(* IEC 61131-3 sources: plc_NativeGateway/src, 67 files *)

(* ---- NG_Add4.st ---- *)
FUNCTION NG_Add4 : DWORD
VAR_INPUT
    a : DWORD;
    b : DWORD;
    c : DWORD;
    d : DWORD;
END_VAR
(* Four uint32 operands fit uint64. A mask implements modulo 2^32 without
   software uint64 division on the AXC F 2152 ARM target. *)
NG_Add4 := TO_DWORD(TO_LWORD(TO_ULINT(a)+TO_ULINT(b)+TO_ULINT(c)+TO_ULINT(d)) AND LWORD#16#FFFFFFFF);
END_FUNCTION

(* ---- NG_Allowed.st ---- *)
FUNCTION NG_Allowed : BOOL
VAR_INPUT
    Parent : INT;
    Keys : NG_Text; (* Delimited with |, including first and last separator. *)
END_VAR
VAR_INPUT
    Doc : NG_Document;
END_VAR
VAR
    i : INT;
    key : STRING[68];
END_VAR
NG_Allowed := FALSE;
IF (Parent < 1) OR (Parent > Doc.Count) THEN RETURN; END_IF;
IF Doc.Tokens[Parent].Kind <> 1 THEN RETURN; END_IF;
i := Parent + 1;
WHILE i < Doc.Tokens[Parent].NextToken DO
    key := CONCAT('|', Doc.Tokens[i].Key, '|');
    IF FIND(Keys,key) = 0 THEN RETURN; END_IF;
    IF Doc.Tokens[i].NextToken <= i THEN RETURN; END_IF;
    i := Doc.Tokens[i].NextToken;
END_WHILE;
NG_Allowed := TRUE;
END_FUNCTION

(* ---- NG_Bool.st ---- *)
FUNCTION NG_Bool : STRING
VAR_INPUT
    Value : BOOL;
END_VAR
IF Value THEN NG_Bool := 'true'; ELSE NG_Bool := 'false'; END_IF;
END_FUNCTION

(* ---- NG_CheckConfig.st ---- *)
FUNCTION NG_CheckConfig : NG_Text
VAR_INPUT
    Config : NG_Config;
END_VAR
VAR
    d : INT;
    p : INT;
    i : INT;
    width : UDINT;
    point : NG_Point;
END_VAR
NG_CheckConfig := 'SCHEMA_INVALID';
IF (Config.PointCount < 0) OR (Config.PointCount > 320) THEN RETURN; END_IF;
IF (Config.DeviceCount < 0) OR (Config.DeviceCount > 50) OR (Config.batchIntervalMs < 1) OR (Config.batchIntervalMs > 86400000) OR (Config.maxBatchPoints < 1) OR (Config.maxBatchPoints > 500) THEN RETURN; END_IF;
FOR d := 1 TO Config.DeviceCount DO
    IF NOT NG_ValidId(Config.Devices[d].deviceId) THEN RETURN; END_IF;
    FOR i := 1 TO d-1 DO
        IF Config.Devices[d].deviceId = Config.Devices[i].deviceId THEN NG_CheckConfig := 'DUPLICATE_DEVICE_ID'; RETURN; END_IF;
    END_FOR;
    IF NOT NG_IPv4(Config.Devices[d].host) THEN NG_CheckConfig := 'BAD_CONFIGURATION'; RETURN; END_IF;
    IF (Config.Devices[d].port = 0) OR (Config.Devices[d].PointCount < 0) OR (Config.Devices[d].PointCount > 32) THEN RETURN; END_IF;
    IF (Config.Devices[d].connectTimeoutMs < 1) OR (Config.Devices[d].connectTimeoutMs > 300000) OR (Config.Devices[d].requestTimeoutMs < 1) OR (Config.Devices[d].requestTimeoutMs > 300000) OR (Config.Devices[d].retryCount > 10) THEN RETURN; END_IF;
    IF (Config.Devices[d].maxReadRegisters > UINT#125) OR (Config.Devices[d].hasMaxRegisterGap AND (Config.Devices[d].maxRegisterGap > UINT#124)) THEN RETURN; END_IF;
    FOR p := 1 TO Config.Devices[d].PointCount DO
        point := Config.Points[Config.Devices[d].PointStart+p-1];
        IF NOT NG_ValidId(point.pointId) THEN RETURN; END_IF;
        FOR i := 1 TO p-1 DO
            IF point.pointId = Config.Points[Config.Devices[d].PointStart+i-1].pointId THEN NG_CheckConfig := 'DUPLICATE_POINT_ID'; RETURN; END_IF;
        END_FOR;
        IF (point.pollIntervalMs < 1) OR (point.pollIntervalMs > 86400000) OR (point.reportIntervalMs < 1) OR (point.reportIntervalMs > 86400000) OR (point.staleAfterMs > 86400000) OR (point.deadband < 0) THEN RETURN; END_IF;
        IF point.staleAfterMs < point.pollIntervalMs THEN NG_CheckConfig := 'INVALID_STALE_INTERVAL'; RETURN; END_IF;
        IF (point.reportMode <> 'cyclic') AND (point.reportMode <> 'change') AND (point.reportMode <> 'change_or_cyclic') THEN RETURN; END_IF;
        IF point.dataType = 'bool' THEN
            width := 1;
            IF (point.area <> 'coil') AND (point.area <> 'discrete_input') THEN RETURN; END_IF;
            IF (point.byteOrder <> '') OR (point.scale <> 1) OR (point.offset <> 0) OR (point.deadband <> 0) THEN RETURN; END_IF;
        ELSE
            IF (point.area <> 'holding_register') AND (point.area <> 'input_register') THEN RETURN; END_IF;
            IF (point.dataType = 'uint16') OR (point.dataType = 'int16') THEN
                width := 1;
                IF (point.byteOrder <> 'AB') AND (point.byteOrder <> 'BA') THEN RETURN; END_IF;
            ELSIF (point.dataType = 'uint32') OR (point.dataType = 'int32') OR (point.dataType = 'float32') THEN
                width := 2;
                IF (point.byteOrder <> 'ABCD') AND (point.byteOrder <> 'BADC') AND (point.byteOrder <> 'CDAB') AND (point.byteOrder <> 'DCBA') THEN RETURN; END_IF;
            ELSE RETURN;
            END_IF;
        END_IF;
        IF TO_UDINT(point.address) + width > 65536 THEN NG_CheckConfig := 'INVALID_ADDRESS'; RETURN; END_IF;
    END_FOR;
END_FOR;
NG_CheckConfig := '';
END_FUNCTION

(* ---- NG_Clip.st ---- *)
FUNCTION NG_Clip : NG_Text
VAR_INPUT
    Value : NG_Text;
END_VAR
IF LEN(Value) > 48 THEN NG_Clip := CONCAT(LEFT(Value,45),'...');
ELSE NG_Clip := Value; END_IF;
END_FUNCTION

(* ---- NG_IPv4.st ---- *)
FUNCTION NG_IPv4 : BOOL
VAR_INPUT
    Host : STRING[253];
END_VAR
VAR
    i : INT;
    dots : INT;
    digits : INT;
    value : INT;
    c : STRING[1];
END_VAR
NG_IPv4 := FALSE; dots := 0; digits := 0; value := 0;
FOR i := 1 TO LEN(Host) DO
    c := MID(Host,1,i);
    IF c = '.' THEN
        IF (digits = 0) OR (value > 255) THEN RETURN; END_IF;
        dots := dots + 1; digits := 0; value := 0;
    ELSIF (c >= '0') AND (c <= '9') THEN
        value := value * 10 + TO_INT(c); digits := digits + 1;
        IF digits > 3 THEN RETURN; END_IF;
    ELSE RETURN;
    END_IF;
END_FOR;
NG_IPv4 := (dots = 3) AND (digits > 0) AND (value <= 255);
END_FUNCTION

(* ---- NG_Member.st ---- *)
FUNCTION NG_Member : INT
VAR_INPUT
    Parent : INT;
    Key : NG_Id;
END_VAR
VAR_INPUT
    Doc : NG_Document;
END_VAR
VAR
    i : INT;
END_VAR
NG_Member := 0;
IF (Parent < 1) OR (Parent > Doc.Count) THEN RETURN; END_IF;
i := Parent + 1;
WHILE i < Doc.Tokens[Parent].NextToken DO
    IF Doc.Tokens[i].Key = Key THEN NG_Member := i; RETURN; END_IF;
    IF Doc.Tokens[i].NextToken <= i THEN RETURN; END_IF;
    i := Doc.Tokens[i].NextToken;
END_WHILE;
END_FUNCTION

(* ---- NG_NumberValid.st ---- *)
FUNCTION NG_NumberValid : BOOL
VAR_INPUT
    s : NG_Text;
END_VAR
VAR
    i : INT;
    n : INT;
    start : INT;
    c : STRING[1];
END_VAR
NG_NumberValid := FALSE;
n := LEN(s); i := 1;
IF n = 0 THEN RETURN; END_IF;
IF MID(s,1,i) = '-' THEN i := i + 1; END_IF;
IF i > n THEN RETURN; END_IF;
c := MID(s,1,i);
IF c = '0' THEN
    i := i + 1;
ELSIF (c >= '1') AND (c <= '9') THEN
    WHILE i <= n DO
        c := MID(s,1,i);
        IF (c < '0') OR (c > '9') THEN EXIT; END_IF;
        i := i + 1;
    END_WHILE;
ELSE RETURN;
END_IF;
IF i > n THEN NG_NumberValid := TRUE; RETURN; END_IF;
IF MID(s,1,i) = '.' THEN
    i := i + 1; start := i;
    WHILE i <= n DO
        c := MID(s,1,i);
        IF (c < '0') OR (c > '9') THEN EXIT; END_IF;
        i := i + 1;
    END_WHILE;
    IF i = start THEN RETURN; END_IF;
END_IF;
IF i > n THEN NG_NumberValid := TRUE; RETURN; END_IF;
c := MID(s,1,i);
IF (c = 'e') OR (c = 'E') THEN
    i := i + 1; IF i > n THEN RETURN; END_IF; c := MID(s,1,i);
    IF (c = '+') OR (c = '-') THEN i := i + 1; END_IF;
    start := i;
    WHILE i <= n DO
        c := MID(s,1,i);
        IF (c < '0') OR (c > '9') THEN EXIT; END_IF;
        i := i + 1;
    END_WHILE;
    IF i = start THEN RETURN; END_IF;
END_IF;
NG_NumberValid := i = n + 1;
END_FUNCTION

(* ---- NG_ProcNumber.st ---- *)
FUNCTION NG_ProcNumber : ULINT
VAR_INPUT
    Text : NG_ProcText;
    Key : STRING[64];
END_VAR
VAR
    p : INT;
    n : INT;
    c : INT;
    started : BOOL;
END_VAR
NG_ProcNumber := 0; started := FALSE; p := FIND(Text,Key); IF p = 0 THEN RETURN; END_IF;
p := p+LEN(Key); n := LEN(Text);
WHILE p <= n DO
    c := GET_CHAR(Text,p);
    IF (c >= 48) AND (c <= 57) THEN NG_ProcNumber := NG_ProcNumber*10+TO_ULINT(c-48); started := TRUE;
    ELSIF started OR ((c <> 32) AND (c <> 9)) THEN RETURN;
    END_IF;
    p := p+1;
END_WHILE;
END_FUNCTION

(* ---- NG_QualityCode.st ---- *)
FUNCTION NG_QualityCode : USINT
VAR_INPUT
    Quality : STRING[24];
END_VAR
NG_QualityCode := 7;
IF Quality='UNKNOWN' THEN NG_QualityCode:=1;
ELSIF Quality='GOOD' THEN NG_QualityCode:=2;
ELSIF Quality='STALE' THEN NG_QualityCode:=3;
ELSIF Quality='BAD_CONNECTION' THEN NG_QualityCode:=4;
ELSIF Quality='BAD_TIMEOUT' THEN NG_QualityCode:=5;
ELSIF Quality='BAD_PROTOCOL' THEN NG_QualityCode:=6;
END_IF;
END_FUNCTION

(* ---- NG_QualityName.st ---- *)
FUNCTION NG_QualityName : NG_Text
VAR_INPUT
    Code : USINT;
END_VAR
CASE Code OF
2: NG_QualityName:='GOOD';
3: NG_QualityName:='STALE';
4: NG_QualityName:='BAD_CONNECTION';
5: NG_QualityName:='BAD_TIMEOUT';
6: NG_QualityName:='BAD_PROTOCOL';
7: NG_QualityName:='BAD_DECODE';
ELSE NG_QualityName:='UNKNOWN';
END_CASE;
END_FUNCTION

(* ---- NG_Quote.st ---- *)
FUNCTION NG_Quote : NG_Quoted
VAR_INPUT
    s : NG_Text;
END_VAR
VAR
    i : INT;
    c : STRING[1];
    character : INT;
    plain : BOOL;
    characters : ARRAY[0..255] OF BYTE;
    copied : BOOL;
    length : INT;
END_VAR
(* Scan once for escaping; common identities take one final concatenation. *)
plain:=TRUE;
length:=LEN(s); copied:=TRUE;
IF length>0 THEN copied:=STRING_COPY(s,characters,UDINT#0,TO_UDINT(length)); END_IF;
FOR i:=1 TO length DO
    IF copied THEN character:=TO_INT(characters[i-1]);
    ELSE character:=GET_CHAR(s,i); END_IF;
    IF (character<32) OR (character=34) OR (character=92) THEN plain:=FALSE; EXIT; END_IF;
END_FOR;
IF plain THEN NG_Quote:=CONCAT('"',s,'"'); RETURN; END_IF;
NG_Quote := '"';
FOR i := 1 TO LEN(s) DO
    c := MID(s,1,i);
    IF c = '"' THEN NG_Quote := CONCAT(NG_Quote,'\\','"');
    ELSIF c = '\\' THEN NG_Quote := CONCAT(NG_Quote,'\\\\');
    ELSIF c = '\n' THEN NG_Quote := CONCAT(NG_Quote,'\\n');
    ELSIF GET_CHAR(c,1) = 13 THEN NG_Quote := CONCAT(NG_Quote,'\\r');
    ELSIF c = '\t' THEN NG_Quote := CONCAT(NG_Quote,'\\t');
    ELSE NG_Quote := CONCAT(NG_Quote,c);
    END_IF;
END_FOR;
NG_Quote := CONCAT(NG_Quote,'"');
END_FUNCTION

(* ---- NG_Range.st ---- *)
FUNCTION NG_Range : BOOL
VAR_INPUT
    Text : NG_Text;
    Minimum : LREAL;
    Maximum : LREAL;
    IntegerOnly : BOOL;
END_VAR
VAR
    n : LREAL;
END_VAR
NG_Range := FALSE;
IF NOT NG_NumberValid(Text) OR (LEN(Text)>20) THEN RETURN; END_IF;
(* UI configuration values do not need exponent notation. *)
IF (FIND(Text,'e')>0) OR (FIND(Text,'E')>0) THEN RETURN; END_IF;
n := TO_LREAL(Text);
NG_Range := (n >= Minimum) AND (n <= Maximum);
IF IntegerOnly AND (n <> TO_LREAL(TO_LINT(n))) THEN NG_Range := FALSE; END_IF;
END_FUNCTION

(* ---- NG_SafeAdd.st ---- *)
FUNCTION NG_SafeAdd : ULINT
VAR_INPUT
    CounterValue : ULINT;
    Delta : ULINT;
END_VAR
IF CounterValue>=ULINT#9007199254740991 THEN NG_SafeAdd:=ULINT#9007199254740991; RETURN; END_IF;
IF Delta>ULINT#9007199254740991-CounterValue THEN
    NG_SafeAdd := ULINT#9007199254740991;
ELSE NG_SafeAdd := CounterValue+Delta;
END_IF;
END_FUNCTION

(* ---- NG_UiJoin.st ---- *)
FUNCTION NG_UiJoin : NG_UiLabel
VAR_INPUT
    A : NG_UiLabel;
    B : NG_UiLabel;
    C : NG_UiLabel;
    D : NG_UiLabel;
    E : NG_UiLabel;
    F : NG_UiLabel;
    G : NG_UiLabel;
    H : NG_UiLabel;
END_VAR
VAR
    Buffer : NG_UiLabel;
    Parts : ARRAY[1..8] OF NG_UiLabel;
    Chunk : NG_UiLabel;
    Remaining : INT;
    i : INT;
END_VAR
(* Explicit intermediates avoid the vendor's default 80-character FU temporary. *)
Parts[1]:=A; Parts[2]:=B; Parts[3]:=C; Parts[4]:=D;
Parts[5]:=E; Parts[6]:=F; Parts[7]:=G; Parts[8]:=H;
Buffer:="";
FOR i:=1 TO 8 DO
    Remaining:=256-LEN(Buffer);
    IF Remaining<=0 THEN EXIT; END_IF;
    Chunk:=Parts[i];
    IF LEN(Chunk)>Remaining THEN Chunk:=LEFT_WSTRING(Chunk,Remaining); END_IF;
    Buffer:=CONCAT_WSTRING(Buffer,Chunk);
END_FOR;
NG_UiJoin:=Buffer;
END_FUNCTION

(* ---- NG_UiText.st ---- *)
FUNCTION NG_UiText : NG_UiLabel
VAR_INPUT
    Value : NG_Text;
    English : BOOL;
END_VAR
NG_UiText:=TO_WSTRING(Value,"");
IF English THEN
IF Value='PERSISTED' THEN NG_UiText:="Saved · no changes";
ELSIF Value='UNSAVED DRAFT' THEN NG_UiText:="Unapplied changes";
ELSIF Value='VERSION CONFLICT' THEN NG_UiText:="Configuration changed";
ELSIF Value='CONNECTED' THEN NG_UiText:="Connected";
ELSIF Value='CONNECTING' THEN NG_UiText:="Connecting";
ELSIF Value='HUB_MANAGED' THEN NG_UiText:="Hub managed";
ELSIF Value='STANDALONE' THEN NG_UiText:="Local maintenance";
ELSIF Value='holding_register' THEN NG_UiText:="Holding register";
ELSIF Value='input_register' THEN NG_UiText:="Input register";
ELSIF Value='discrete_input' THEN NG_UiText:="Discrete input";
ELSIF Value='cyclic' THEN NG_UiText:="Cyclic";
ELSIF Value='change' THEN NG_UiText:="On change";
ELSIF Value='change_or_cyclic' THEN NG_UiText:="Change or cyclic";
ELSIF Value='Startup identity persisted; MQTT starting.' THEN NG_UiText:="Saved configuration restored automatically. No need to save again.";
ELSIF Value='true' THEN NG_UiText:="Enabled";
ELSIF Value='TRUE' THEN NG_UiText:="Enabled";
ELSIF Value='false' THEN NG_UiText:="Disabled";
ELSIF Value='FALSE' THEN NG_UiText:="Disabled";
ELSIF Value='HUB_MANAGED - local device/point changes blocked' THEN NG_UiText:="Managed by Hub: edit and publish devices, points and periods in Hub. Connection maintenance is available here.";
ELSIF Value='STANDALONE - local maintenance enabled' THEN NG_UiText:="Standalone: edit devices and points → save to draft → review and activate.";
END_IF;
RETURN;
END_IF;
IF Value='Open the management mode confirmation before saving.' THEN NG_UiText:="请先打开模式切换确认页，检查选项后再确认。";
ELSIF Value='Waiting for initial Hub configuration. Existing local acquisition is retained.' THEN NG_UiText:="正在等待平台首次配置；现有本地采集保留，暂不向平台上报。";
ELSIF Value='Invalid management mode.' THEN NG_UiText:="管理模式无效，请重新选择平台管理或本地维护。";
ELSIF Value='MAINTENANCE - incoming platform configuration locked' THEN NG_UiText:="本地维护：平台配置暂不应用；修改后请交还平台，避免两端配置冲突。";
ELSIF Value='Hub owns configuration. Local maintenance requires manual confirmation.' THEN NG_UiText:="当前由平台管理。需要本地编辑时，请手动进入维护。";
ELSIF Value='Local changes active. Acquisition continues; Hub data reporting is paused.' THEN NG_UiText:="本地改动已生效：继续采集，暂停写入平台；交还时恢复平台配置。";
ELSIF Value='Local maintenance active. Hub configuration is locked until you return ownership.' THEN NG_UiText:="本地维护中：平台配置暂不应用。维护完成后请交还平台。";
ELSIF Value='The selected management mode is already active.' THEN NG_UiText:="已处于所选模式，无需重复切换。";
ELSIF Value='Saving management mode; existing identity is retained.' THEN NG_UiText:="正在保存管理模式，保留当前网关标识。";
ELSIF Value='Management mode saved. Check the ownership guidance above.' THEN NG_UiText:="管理模式已保存并生效，请查看上方的管理说明。";
ELSIF Value='Clearing local configuration and version baseline...' THEN NG_UiText:="正在清空本地点表与版本基线，请稍候。";
ELSIF Value='Open the reset confirmation before clearing local configuration.' THEN NG_UiText:="请先打开重置确认页后再确认清空。";
ELSIF Value='Local configuration and version baseline cleared; requesting fresh config from Hub.' THEN NG_UiText:="已清空本地点表与版本基线，正在重连并向平台重新拉取配置。";
ELSIF Value='Check broker URI, gateway ID, client ID and time zone.' THEN NG_UiText:="请检查服务器地址、网关标识与时区。";
ELSIF Value='Broker settings saved; configuration ownership is unchanged.' THEN NG_UiText:="连接设置已保存，正在重连；管理模式保持不变。";
ELSIF Value='CONNECTED' THEN NG_UiText:="已连接";
ELSIF Value='CONNECTING' THEN NG_UiText:="正在连接";
ELSIF Value='ONLINE' THEN NG_UiText:="在线";
ELSIF Value='OFFLINE' THEN NG_UiText:="离线";
ELSIF Value='DEGRADED' THEN NG_UiText:="部分异常";
ELSIF Value='DISABLED' THEN NG_UiText:="已停用";
ELSIF Value='UNCONFIGURED' THEN NG_UiText:="未配置";
ELSIF Value='DRAFT' THEN NG_UiText:="待生效";
ELSIF Value='GOOD' THEN NG_UiText:="正常";
ELSIF Value='BAD' THEN NG_UiText:="异常";
ELSIF Value='STALE' THEN NG_UiText:="已过期";
ELSIF Value='UNKNOWN' THEN NG_UiText:="暂无数据";
ELSIF Value='BAD_COMMUNICATION' THEN NG_UiText:="通信异常";
ELSIF Value='BAD_CONFIGURATION' THEN NG_UiText:="配置有误";
ELSIF Value='true' THEN NG_UiText:="启用";
ELSIF Value='TRUE' THEN NG_UiText:="启用";
ELSIF Value='false' THEN NG_UiText:="停用";
ELSIF Value='FALSE' THEN NG_UiText:="停用";
ELSIF Value='PERSISTED' THEN NG_UiText:="已保存，无待生效修改";
ELSIF Value='UNSAVED DRAFT' THEN NG_UiText:="有待生效的修改";
ELSIF Value='VERSION CONFLICT' THEN NG_UiText:="配置已变更，请放弃旧草稿";
ELSIF Value='HUB_MANAGED' THEN NG_UiText:="平台统一管理";
ELSIF Value='STANDALONE' THEN NG_UiText:="本地维护";
ELSIF Value='HUB_MANAGED - local device/point changes blocked' THEN NG_UiText:="平台管理：在 Hub 编辑设备、点位与周期并发布；此处查看和维护连接。";
ELSIF Value='STANDALONE - local maintenance enabled' THEN NG_UiText:="本地管理：编辑设备和点位 → 保存到待生效配置 → 确认生效并保存。";
ELSIF Value='holding_register' THEN NG_UiText:="保持寄存器";
ELSIF Value='input_register' THEN NG_UiText:="输入寄存器";
ELSIF Value='coil' THEN NG_UiText:="线圈";
ELSIF Value='discrete_input' THEN NG_UiText:="离散输入";
ELSIF Value='cyclic' THEN NG_UiText:="定时上报";
ELSIF Value='change' THEN NG_UiText:="变化时上报";
ELSIF Value='change_or_cyclic' THEN NG_UiText:="变化或定时上报";
ELSIF Value='voltage' THEN NG_UiText:="电压";
ELSIF Value='current' THEN NG_UiText:="电流";
ELSIF Value='frequency' THEN NG_UiText:="频率";
ELSIF Value='power' THEN NG_UiText:="功率";
ELSIF Value='energy' THEN NG_UiText:="累计电能";
ELSIF Value='No device selected' THEN NG_UiText:="暂无设备，请先添加设备";
ELSIF Value='No point selected' THEN NG_UiText:="暂无点位，请先添加点位";
ELSIF Value='HUB_MANAGED: publish device and point changes from Hub.' THEN NG_UiText:="当前由平台管理，请在 Hub 修改并发布设备和点位配置。";
ELSIF Value='Display refreshed from active configuration. Unapplied draft discarded.' THEN NG_UiText:="已按当前运行配置更新显示，未生效的草稿已放弃。";
ELSIF Value='Loaded persisted active configuration.' THEN NG_UiText:="已按控制器当前运行配置更新显示。";
ELSIF Value='Capacity reached: 50 devices.' THEN NG_UiText:="设备数量已达上限：50 台。";
ELSIF Value='Capacity reached: 32 points/device, 320 shared points.' THEN NG_UiText:="点位数量已达上限：每台 32 个，总计 320 个。";
ELSIF Value='New device: save into draft, then add its points.' THEN NG_UiText:="填写连接参数并保存设备，再为该设备添加点位。";
ELSIF Value='Save a device into the draft first.' THEN NG_UiText:="请先保存设备，再添加该设备的点位。";
ELSIF Value='New point: save into draft, then apply the complete draft.' THEN NG_UiText:="填写寄存器与周期，保存点位后再确认配置生效。";
ELSIF Value='Busy: configuration transaction in progress. Try again shortly.' THEN NG_UiText:="正在保存配置，请稍候再试。";
ELSIF Value='Device index 1..50; point index 1..32.' THEN NG_UiText:="请检查设备序号（1～50）和点位序号（1～32）。";
ELSIF Value='Invalid device fields: check ID, name, IPv4, port and timeout values.' THEN NG_UiText:="设备未保存：检查唯一标识、名称、地址、端口与超时。";
ELSIF Value='Device saved to draft. Apply draft to persist.' THEN NG_UiText:="设备已加入待生效配置。检查点位后，点击“使配置生效”。";
ELSIF Value='Invalid point fields; save the device first and check numeric fields.' THEN NG_UiText:="点位未保存：先保存设备，再检查地址、周期、倍率等数值。";
ELSIF Value='Point saved to draft. Apply draft to persist.' THEN NG_UiText:="点位已加入待生效配置。点击“使配置生效”后开始使用。";
ELSIF Value='Device and points removed from draft. Apply to persist.' THEN NG_UiText:="设备及其点位已从草稿移除，确认配置生效后才停止采集。";
ELSIF Value='Point removed from draft. Apply to persist.' THEN NG_UiText:="点位已从草稿移除，确认配置生效后才停止采集。";
ELSIF Value='Invalid device polling/report period.' THEN NG_UiText:="周期未修改：采集与上报周期必须为有效的毫秒数。";
ELSIF Value='Device point periods updated in draft. Apply to persist.' THEN NG_UiText:="该设备的点位周期已加入待生效配置，请确认生效。";
ELSIF Value='VERSION_CONFLICT: reload active configuration before applying.' THEN NG_UiText:="运行配置已有更新。请放弃旧草稿，按最新配置重新编辑。";
ELSIF Value='Invalid gateway batch settings.' THEN NG_UiText:="请检查组批周期与每包点数（1～64）。";
ELSIF Value='Saving, hashing and reading back configuration...' THEN NG_UiText:="正在保存并校验配置，请稍候。";
ELSIF Value='Check broker/mode/ID. Mode change requires a new Gateway ID to isolate configuration history.' THEN NG_UiText:="连接未保存：检查地址、网关标识、客户端标识与模式；换模式须换网关标识。";
ELSIF Value='Saving broker settings...' THEN NG_UiText:="正在保存消息服务器连接设置，请稍候。";
ELSIF Value='APPLIED: configuration saved and activated.' THEN NG_UiText:="配置已生效并保存；重启后将自动恢复。";
ELSIF Value='Broker/mode saved; identity changes reset local baseline.' THEN NG_UiText:="连接设置已保存，正在自动重连；新身份需由平台重新下发配置。";
ELSIF Value='Startup identity persisted; MQTT starting.' THEN NG_UiText:="已自动恢复保存的配置，无需重复保存。";
ELSIF Value='Persisting unique startup identity before MQTT...' THEN NG_UiText:="正在保存启动信息，随后自动连接消息服务器。";
ELSIF Value='STORAGE_ERROR: active configuration unchanged.' THEN NG_UiText:="保存失败，运行配置保持原样。请检查控制器存储。";
ELSIF Value='Saving / validating durable file...' THEN NG_UiText:="正在写入并校验控制器配置文件……";
ELSIF Value='STORAGE ERROR: configuration not committed.' THEN NG_UiText:="配置保存失败，请检查控制器存储。";
ELSIF Value='Restoring saved configuration...' THEN NG_UiText:="正在恢复已保存配置，随后自动连接并采集。";
ELSIF Value='Broker unavailable. Retrying automatically; local acquisition continues.' THEN NG_UiText:="消息服务器暂不可用，正在自动重连；本地采集继续运行。";
ELSIF Value='MQTT_DISCONNECTED' THEN NG_UiText:="连接中断，自动重连中";
ELSIF Value='MQTT_CONNECT_ERROR' THEN NG_UiText:="连接失败，自动重试中";
ELSIF Value='MQTT_TIMEOUT' THEN NG_UiText:="连接超时，自动重试中";
ELSIF Value='MQTT_PUBLISH_ERROR' THEN NG_UiText:="发送失败，自动重连中";
ELSIF Value='MQTT_CLIENT_ERROR' THEN NG_UiText:="通信组件异常，自动重试中";
ELSIF Value='MQTT_SUBSCRIBE_ERROR' THEN NG_UiText:="订阅失败，自动重试中";
ELSIF Value='MQTT_CONSUME_ERROR' THEN NG_UiText:="接收失败，自动重试中";
ELSIF Value='SCHEMA_INVALID' THEN NG_UiText:="配置格式或取值不正确，请检查点位详情。";
ELSIF Value='DUPLICATE_DEVICE_ID' THEN NG_UiText:="设备标识重复，请使用唯一标识。";
ELSIF Value='DUPLICATE_POINT_ID' THEN NG_UiText:="同一设备内点位标识重复。";
ELSIF Value='INVALID_STALE_INTERVAL' THEN NG_UiText:="过期时间必须不小于采集周期。";
ELSIF Value='INVALID_ADDRESS' THEN NG_UiText:="寄存器地址范围无效。";
ELSIF Value='BAD_CONNECTION' THEN NG_UiText:="连接异常";
ELSIF Value='BAD_TIMEOUT' THEN NG_UiText:="请求超时";
ELSIF Value='BAD_PROTOCOL' THEN NG_UiText:="报文异常";
ELSIF Value='BAD_DECODE' THEN NG_UiText:="数据解码异常";
END_IF;
END_FUNCTION

(* ---- NG_Unix.st ---- *)
FUNCTION NG_Unix : ULINT
VAR_INPUT
    Clock : RTC_TYPE;
    UtcOffsetMinutes : INT;
END_VAR
VAR
    y : DINT;
    m : DINT;
    days : LINT;
    md : DINT;
    seconds : LINT;
END_VAR
NG_Unix := 0;
IF (Clock.YEAR < 2020) OR (Clock.YEAR > 2199) OR (Clock.MONTH < 1) OR (Clock.MONTH > 12) OR (Clock.DAY < 1) OR (Clock.DAY > 31) THEN RETURN; END_IF;
days := 0;
FOR y := 1970 TO TO_DINT(Clock.YEAR)-1 DO
    days := days + 365;
    IF ((y MOD 4 = 0) AND (y MOD 100 <> 0)) OR (y MOD 400 = 0) THEN days := days + 1; END_IF;
END_FOR;
FOR m := 1 TO TO_DINT(Clock.MONTH)-1 DO
    CASE m OF
        4,6,9,11: md := 30;
        2:
            md := 28; y := TO_DINT(Clock.YEAR);
            IF ((y MOD 4 = 0) AND (y MOD 100 <> 0)) OR (y MOD 400 = 0) THEN md := 29; END_IF;
        ELSE md := 31;
    END_CASE;
    days := days + md;
END_FOR;
days := days + Clock.DAY - 1;
seconds := days * 86400 + TO_LINT(Clock.HOURS) * 3600 + TO_LINT(Clock.MINUTES) * 60 + Clock.SECONDS - TO_LINT(UtcOffsetMinutes)*60;
IF seconds > 0 THEN NG_Unix := TO_ULINT(seconds)*1000; END_IF;
END_FUNCTION

(* ---- NG_ValidId.st ---- *)
FUNCTION NG_ValidId : BOOL
VAR_INPUT
    s : NG_Id;
END_VAR
VAR
    i : INT;
    c : STRING[1];
END_VAR
NG_ValidId := (LEN(s) > 0) AND (LEN(s) <= 64);
FOR i := 1 TO LEN(s) DO
    c := MID(s, 1, i);
    IF NOT (((c >= 'A') AND (c <= 'Z')) OR ((c >= 'a') AND (c <= 'z')) OR ((c >= '0') AND (c <= '9')) OR ((i > 1) AND ((c = '.') OR (c = '_') OR (c = '-')))) THEN
        NG_ValidId := FALSE;
    END_IF;
END_FOR;
END_FUNCTION

(* ---- NG_WireCode.st ---- *)
FUNCTION NG_WireCode : NG_Text
VAR_INPUT
    Code : NG_Text;
    IsPatch : BOOL;
END_VAR
IF FIND('|SCHEMA_INVALID|INVALID_JSON|PAYLOAD_TOO_LARGE|GATEWAY_MISMATCH|DUPLICATE_DEVICE_ID|DUPLICATE_POINT_ID|DUPLICATE_NODE_ID|INVALID_ADDRESS|INVALID_STALE_INTERVAL|POINT_LIMIT_EXCEEDED|VERSION_CONFLICT|STALE_VERSION|RESOURCE_LIMIT|STORAGE_ERROR|APPLY_FAILED|UNKNOWN_CONFIG_VERSION|UNKNOWN_DEVICE|UNKNOWN_POINT|EXPIRED_DATA|INVALID_TIMESTAMP|DUPLICATE_VALUE|',CONCAT('|',Code,'|')) > 0 THEN NG_WireCode := Code;
ELSIF IsPatch AND (Code = 'RETAINED_PATCH') THEN NG_WireCode := 'OPERATION_CONFLICT';
ELSIF IsPatch AND (FIND('|BASE_CONFIG_MISMATCH|DEVICE_EXISTS|DEVICE_NOT_FOUND|OPERATION_CONFLICT|',CONCAT('|',Code,'|'))>0) THEN NG_WireCode := Code;
ELSE NG_WireCode := 'APPLY_FAILED';
END_IF;
END_FUNCTION

(* ---- NG_AckFields.st ---- *)
FUNCTION_BLOCK NG_AckFields
VAR_INPUT
    Parent : INT;
    ErrorObject : BOOL;
END_VAR
VAR_IN_OUT
    Doc : NG_Document;
END_VAR
VAR_OUTPUT
    Valid : BOOL;
    Fields : ARRAY[1..6] OF INT;
END_VAR
VAR
    i : INT;
    j : INT;
    field : INT;
    count : INT;
END_VAR
(* A bounded, reference-based index for the two ACK object shapes. It keeps
   the full document out of FUNCTION VAR_INPUT argument copies. *)
Valid:=FALSE; FOR j:=1 TO 6 DO Fields[j]:=0; END_FOR;
IF (Parent<1) OR (Parent>Doc.Count) THEN RETURN; END_IF;
IF Doc.Tokens[Parent].Kind<>1 THEN RETURN; END_IF;
i:=Parent+1; count:=0;
WHILE i<Doc.Tokens[Parent].NextToken DO
    count:=count+1; IF count>6 THEN RETURN; END_IF;
    IF (i>Doc.Count) OR (i>8192) THEN RETURN; END_IF;
    field:=0;
    IF ErrorObject THEN
        IF Doc.Tokens[i].Key='code' THEN field:=1;
        ELSIF Doc.Tokens[i].Key='path' THEN field:=2;
        ELSIF Doc.Tokens[i].Key='message' THEN field:=3;
        ELSIF Doc.Tokens[i].Key='deviceId' THEN field:=4;
        ELSIF Doc.Tokens[i].Key='pointId' THEN field:=5; END_IF;
    ELSE
        IF Doc.Tokens[i].Key='schemaVersion' THEN field:=1;
        ELSIF Doc.Tokens[i].Key='gatewayId' THEN field:=2;
        ELSIF Doc.Tokens[i].Key='timestamp' THEN field:=3;
        ELSIF Doc.Tokens[i].Key='messageId' THEN field:=4;
        ELSIF Doc.Tokens[i].Key='status' THEN field:=5;
        ELSIF Doc.Tokens[i].Key='errors' THEN field:=6; END_IF;
    END_IF;
    IF field=0 THEN RETURN; END_IF;
    IF Fields[field]<>0 THEN RETURN; END_IF;
    Fields[field]:=i;
    IF (Doc.Tokens[i].NextToken<=i) OR (Doc.Tokens[i].NextToken>Doc.Tokens[Parent].NextToken) THEN RETURN; END_IF;
    i:=Doc.Tokens[i].NextToken;
END_WHILE;
IF i<>Doc.Tokens[Parent].NextToken THEN RETURN; END_IF;
IF ErrorObject THEN
    IF (Fields[1]=0) OR (Fields[2]=0) OR (Fields[3]=0) THEN RETURN; END_IF;
ELSE
    FOR j:=1 TO 6 DO IF Fields[j]=0 THEN RETURN; END_IF; END_FOR;
END_IF;
Valid:=TRUE;
END_FUNCTION_BLOCK

(* ---- NG_AuditAssociation.st ---- *)
FUNCTION_BLOCK NG_AuditAssociation
VAR_INPUT
    Slot : UINT;
    MessageId : NG_Id;
END_VAR
VAR_IN_OUT
    Buffer : NG_Buffer;
END_VAR
VAR
    index : UINT;
    configSlot : UINT;
    j : UINT;
    offset : UINT;
END_VAR
IF NOT Buffer.AuditEnabled THEN RETURN; END_IF;
IF (Slot<1) OR (Slot>16) THEN Buffer.CaptureStopped:=TRUE; Buffer.EvidenceComplete:=FALSE; RETURN; END_IF;
IF Buffer.AssociationWriteSeq>=ULINT#9007199254740991 THEN Buffer.CaptureStopped:=TRUE; RETURN; END_IF;
IF Buffer.AssociationWriteSeq-Buffer.AssociationReadSeq>=32 THEN
    index:=TO_UINT(Buffer.AssociationReadSeq MOD 32)+1;
    configSlot:=Buffer.Associations[index].ConfigSlot;
    IF (configSlot<1) OR (configSlot>4) THEN Buffer.CaptureStopped:=TRUE; Buffer.EvidenceComplete:=FALSE; RETURN; END_IF;
    IF Buffer.Configs[configSlot].References=0 THEN Buffer.CaptureStopped:=TRUE; Buffer.EvidenceComplete:=FALSE; RETURN; END_IF;
    Buffer.Configs[configSlot].References:=Buffer.Configs[configSlot].References-1;
    Buffer.AssociationReadSeq:=Buffer.AssociationReadSeq+1;
    Buffer.AssociationDropped:=NG_SafeAdd(Buffer.AssociationDropped,ULINT#1); Buffer.EvidenceComplete:=FALSE;
END_IF;
Buffer.AssociationWriteSeq:=Buffer.AssociationWriteSeq+1; index:=TO_UINT((Buffer.AssociationWriteSeq-1) MOD 32)+1;
configSlot:=Buffer.BatchOwners[Slot].ConfigSlot;
IF (configSlot<1) OR (configSlot>4) THEN Buffer.CaptureStopped:=TRUE; Buffer.EvidenceComplete:=FALSE; RETURN; END_IF;
Buffer.Associations[index].Ordinal:=Buffer.AssociationWriteSeq;
Buffer.Associations[index].MessageId:=MessageId; Buffer.Associations[index].Digest:=Buffer.BatchOwners[Slot].Digest;
Buffer.Associations[index].ConfigSlot:=configSlot; Buffer.Associations[index].ConfigGeneration:=Buffer.Configs[configSlot].Generation;
Buffer.Associations[index].BatchGeneration:=Buffer.BatchGenerations[Slot]; Buffer.Associations[index].Category:=Buffer.BatchOwners[Slot].Category;
Buffer.Associations[index].Count:=Buffer.BatchOwners[Slot].Count; offset:=(Slot-1)*64;
FOR j:=1 TO Buffer.BatchOwners[Slot].Count DO Buffer.Associations[index].SampleSeqs[j]:=Buffer.Records[Buffer.BatchRefs[offset+j]].SampleSeq; END_FOR;
Buffer.Configs[configSlot].References:=Buffer.Configs[configSlot].References+1;
END_FUNCTION_BLOCK

(* ---- NG_AuditCapture.st ---- *)
FUNCTION_BLOCK NG_AuditCapture
VAR_IN_OUT
    Buffer : NG_Buffer;
    Event : NG_CaptureEvent;
END_VAR
VAR
    index : UINT;
    oldIndex : UINT;
    configSlot : UINT;
END_VAR

IF NOT Buffer.AuditEnabled THEN RETURN; END_IF;
IF (Event.SampleSeq=0) OR (Event.ConfigSlot<1) OR (Event.ConfigSlot>4) THEN
    Buffer.CaptureStopped:=TRUE; Buffer.EvidenceComplete:=FALSE; RETURN;
END_IF;
IF Buffer.AuditWriteSeq-Buffer.AuditReadSeq>=512 THEN
    oldIndex:=TO_UINT(Buffer.AuditReadSeq MOD 512)+1;
    configSlot:=Buffer.AuditEvents[oldIndex].Event.ConfigSlot;
    IF (configSlot<1) OR (configSlot>4) THEN Buffer.CaptureStopped:=TRUE; Buffer.EvidenceComplete:=FALSE; RETURN; END_IF;
    IF Buffer.Configs[configSlot].References=0 THEN Buffer.CaptureStopped:=TRUE; Buffer.EvidenceComplete:=FALSE; RETURN; END_IF;
    Buffer.Configs[configSlot].References:=Buffer.Configs[configSlot].References-1;
    Buffer.AuditReadSeq:=Buffer.AuditReadSeq+1;
    Buffer.AuditDropped:=NG_SafeAdd(Buffer.AuditDropped,ULINT#1); Buffer.EvidenceComplete:=FALSE;
END_IF;
index:=TO_UINT((Event.SampleSeq-1) MOD 512)+1;
Buffer.AuditEvents[index].Event:=Event; Buffer.AuditEvents[index].Decision:=0; Buffer.AuditEvents[index].Reason:=0;
Buffer.Configs[Event.ConfigSlot].References:=Buffer.Configs[Event.ConfigSlot].References+1;
Buffer.AuditWriteSeq:=Event.SampleSeq;
END_FUNCTION_BLOCK

(* ---- NG_AuditDecision.st ---- *)
FUNCTION_BLOCK NG_AuditDecision
VAR_INPUT
    SampleSeq : ULINT;
    Decision : USINT;
    Reason : USINT;
END_VAR
VAR_IN_OUT
    Buffer : NG_Buffer;
END_VAR
VAR
    index : UINT;
END_VAR

IF NOT Buffer.AuditEnabled OR (SampleSeq=0) THEN RETURN; END_IF;
index:=TO_UINT((SampleSeq-1) MOD 512)+1;
IF (SampleSeq>Buffer.AuditReadSeq) AND (Buffer.AuditEvents[index].Event.SampleSeq=SampleSeq) THEN
    Buffer.AuditEvents[index].Decision:=Decision; Buffer.AuditEvents[index].Reason:=Reason;
ELSE Buffer.EvidenceComplete:=FALSE;
END_IF;
END_FUNCTION_BLOCK

(* ---- NG_AuditDrain.st ---- *)
FUNCTION_BLOCK NG_AuditDrain
VAR_INPUT
    BootId : NG_Id;
END_VAR
VAR_IN_OUT
    Buffer : NG_Buffer;
END_VAR
VAR
    index : UINT;
    configSlot : UINT;
    n : INT;
END_VAR
IF (Buffer.AuditAckBootId=BootId) AND (Buffer.AuditAckSeq<=Buffer.AuditWriteSeq) THEN
    FOR n:=1 TO 8 DO
        IF Buffer.AuditReadSeq>=Buffer.AuditAckSeq THEN EXIT; END_IF;
        index:=TO_UINT(Buffer.AuditReadSeq MOD 512)+1;
        IF Buffer.AuditEvents[index].Event.SampleSeq<>Buffer.AuditReadSeq+1 THEN Buffer.EvidenceComplete:=FALSE; RETURN; END_IF;
        IF Buffer.AuditEvents[index].Decision=0 THEN EXIT; END_IF;
        configSlot:=Buffer.AuditEvents[index].Event.ConfigSlot;
        IF (configSlot<1) OR (configSlot>4) THEN Buffer.EvidenceComplete:=FALSE; RETURN; END_IF;
        IF Buffer.Configs[configSlot].References=0 THEN Buffer.EvidenceComplete:=FALSE; RETURN; END_IF;
        Buffer.Configs[configSlot].References:=Buffer.Configs[configSlot].References-1;
        Buffer.AuditReadSeq:=Buffer.AuditReadSeq+1;
    END_FOR;
END_IF;
IF (Buffer.AssociationAckBootId=BootId) AND (Buffer.AssociationAckSeq<=Buffer.AssociationWriteSeq) THEN
    FOR n:=1 TO 4 DO
        IF Buffer.AssociationReadSeq>=Buffer.AssociationAckSeq THEN EXIT; END_IF;
        index:=TO_UINT(Buffer.AssociationReadSeq MOD 32)+1;
        IF Buffer.Associations[index].Ordinal<>Buffer.AssociationReadSeq+1 THEN Buffer.EvidenceComplete:=FALSE; RETURN; END_IF;
        configSlot:=Buffer.Associations[index].ConfigSlot;
        IF (configSlot<1) OR (configSlot>4) THEN Buffer.EvidenceComplete:=FALSE; RETURN; END_IF;
        IF Buffer.Configs[configSlot].References=0 THEN Buffer.EvidenceComplete:=FALSE; RETURN; END_IF;
        Buffer.Configs[configSlot].References:=Buffer.Configs[configSlot].References-1;
        Buffer.AssociationReadSeq:=Buffer.AssociationReadSeq+1;
    END_FOR;
END_IF;
END_FUNCTION_BLOCK

(* ---- NG_BatchBuilder.st ---- *)
FUNCTION_BLOCK NG_BatchBuilder
VAR_INPUT
    GateOpen : BOOL;
    NowMs : ULINT;
    UnixMs : ULINT;
    GatewayId : NG_Id;
    BootId : NG_Id;
    BatchIntervalMs : UDINT;
END_VAR
VAR_IN_OUT
    Buffer : NG_Buffer;
    Packets : ARRAY[1..16] OF NG_Packet;
    Sequence : ULINT;
END_VAR
VAR_OUTPUT
    Busy : BOOL;
END_VAR
VAR
    Digest : NG_StringSHA256;
    Audit : NG_AuditAssociation;
    Stage : UINT;
    Slot : UINT;
    ConfigSlot : UINT;
    Category : UINT;
    q : UINT;
    r : UINT;
    j : UINT;
    offset : UINT;
    countHistory : UINT;
    countNew : UINT;
    n : INT;
    d : INT;
    deviceId : NG_Id;
    valueJson : STRING[80];
    item : STRING[1024];
    bytesNeeded : INT;
    duplicate : BOOL;
    finish : BOOL;
    lastStart : ULINT;
    first : BOOL := TRUE;
    MaterialClockRevision : ULINT;
    windowOpen : BOOL;
    generation : UDINT;
    seenEpoch : UDINT;
    seenPointEpoch : ARRAY[1..320] OF UDINT;
    pointIndex : UINT;
    HeaderUnixMs : ULINT;
    HeaderSequence : ULINT;
    DeviceQuoteSlot : UINT;
    DeviceQuoteGeneration : UDINT;
    DeviceQuoteEpoch : UDINT;
    DeviceQuoteSeen : ARRAY[1..50] OF UDINT;
    DeviceQuotes : ARRAY[1..50] OF STRING[132];
    QuotedDevice : STRING[132];
    ItemPhase : USINT;
    ItemRecord : UINT;
    ItemGeneration : UDINT;
    CachedUtc : ULINT;
    CachedUtcText : STRING[32];
    CachedQuality : USINT;
    CachedQualityText : STRING[40];
    HaveUtc : BOOL;
    HaveQuality : BOOL;
END_VAR
Busy:=Stage<>0;
IF Stage<>0 THEN
    IF (Buffer.BatchGenerations[Slot]<>generation) OR (Buffer.BatchOwners[Slot].State<>1) THEN Stage:=0; END_IF;
END_IF;
IF (Stage<>0) AND (NOT GateOpen OR (Buffer.PlatformTime AND (MaterialClockRevision<>Buffer.ClockRevision))) THEN
    Category:=TO_UINT(Buffer.BatchOwners[Slot].Category); offset:=(Slot-1)*64;
    FOR n:=TO_INT(Buffer.BatchOwners[Slot].Count) TO 1 BY -1 DO
        r:=Buffer.BatchRefs[offset+TO_UINT(n)];
        Buffer.RecordStates[r]:=1; Buffer.FreeSlots[r]:=Buffer.QueueHead[Category];
        Buffer.QueueHead[Category]:=r; IF Buffer.QueueTail[Category]=0 THEN Buffer.QueueTail[Category]:=r; END_IF;
        Buffer.BatchRefs[offset+TO_UINT(n)]:=0;
    END_FOR;
    Buffer.BatchOwners[Slot].State:=0; Buffer.BatchOwners[Slot].Count:=0;
    Packets[Slot].MessageId:=''; Packets[Slot].Payload:=''; Stage:=0;
END_IF;
IF Stage=0 THEN
    IF Buffer.WorkDeadlineUs>0 THEN IF GET_MICROSECONDS(TRUE)+ULINT#180>=Buffer.WorkDeadlineUs THEN RETURN; END_IF; END_IF;
    Digest(Execute:=FALSE,Length:=UDINT#0,Payload:=Packets[1].Payload);
    Busy:=FALSE;
    IF (Buffer.QueueHead[1]=0) AND (Buffer.QueueHead[2]=0) THEN windowOpen:=FALSE; END_IF;
    IF NOT GateOpen OR (UnixMs=0) OR (NOT windowOpen AND NOT first AND (NowMs<lastStart+TO_ULINT(BatchIntervalMs))) THEN RETURN; END_IF;
    countHistory:=0; countNew:=0; Slot:=0;
    FOR q:=1 TO 16 DO
        IF Buffer.BatchOwners[q].State=0 THEN IF Slot=0 THEN Slot:=q; END_IF;
        ELSIF Buffer.BatchOwners[q].State<>3 THEN
            IF Buffer.BatchOwners[q].Category=1 THEN countHistory:=countHistory+1; ELSE countNew:=countNew+1; END_IF;
        END_IF;
    END_FOR;
    IF Slot=0 THEN RETURN; END_IF;
    Category:=TO_UINT(Buffer.PreferMaterialize);
    IF ((Category=1) AND ((Buffer.QueueHead[1]=0) OR (countHistory>=7))) OR
       ((Category=2) AND ((Buffer.QueueHead[2]=0) OR (countNew>=7))) THEN Category:=UINT#3-Category; END_IF;
    IF ((Category=1) AND ((Buffer.QueueHead[1]=0) OR (countHistory>=7))) OR
       ((Category=2) AND ((Buffer.QueueHead[2]=0) OR (countNew>=7))) THEN RETURN; END_IF;
    r:=Buffer.QueueHead[Category]; ConfigSlot:=Buffer.Records[r].ConfigSlot;
    IF (Buffer.Configs[ConfigSlot].GatewayId<>GatewayId) OR (Buffer.Configs[ConfigSlot].CaptureBootId<>BootId) THEN RETURN; END_IF;
    (* Lazy bounded quote cache follows the pinned dictionary's slot AND generation.
       NG_Id has at most 64 characters; escaped JSON needs at most 130 characters. *)
    IF (DeviceQuoteSlot<>ConfigSlot) OR (DeviceQuoteGeneration<>Buffer.Configs[ConfigSlot].Generation) THEN
        IF DeviceQuoteEpoch=UDINT#4294967295 THEN Buffer.CaptureStopped:=TRUE; RETURN; END_IF;
        DeviceQuoteEpoch:=DeviceQuoteEpoch+1;
        DeviceQuoteSlot:=ConfigSlot; DeviceQuoteGeneration:=Buffer.Configs[ConfigSlot].Generation;
    END_IF;
    IF (Sequence>=ULINT#9007199254740991) OR (Buffer.BatchGenerations[Slot]=UDINT#4294967295) THEN Buffer.CaptureStopped:=TRUE; RETURN; END_IF;
    IF seenEpoch=UDINT#4294967295 THEN Buffer.CaptureStopped:=TRUE; RETURN; END_IF;
    seenEpoch:=seenEpoch+1;
    Sequence:=Sequence+1; Buffer.BatchGenerations[Slot]:=Buffer.BatchGenerations[Slot]+1; generation:=Buffer.BatchGenerations[Slot];
    Packets[Slot].MessageId:=CONCAT('d-',BootId,'-',TO_STRING(Sequence,'{0:d}'));
    IF LEN(Packets[Slot].MessageId)>64 THEN Buffer.CaptureStopped:=TRUE; RETURN; END_IF;
    (* Freeze envelope values at reservation; quoting is split into bounded steps. *)
    HeaderUnixMs:=UnixMs; HeaderSequence:=Sequence; MaterialClockRevision:=Buffer.ClockRevision;
    Packets[Slot].Payload:='';
    Packets[Slot].WasSent:=FALSE; Packets[Slot].Attempts:=0; Packets[Slot].Dead:=FALSE;
    Packets[Slot].LastSentMs:=0; Packets[Slot].RetryAtMs:=0; Packets[Slot].LastError:='';
    Buffer.BatchOwners[Slot].State:=1; Buffer.BatchOwners[Slot].Count:=0;
    Buffer.BatchOwners[Slot].Category:=TO_USINT(Category); Buffer.BatchOwners[Slot].ConfigSlot:=ConfigSlot;
    Buffer.BatchOwners[Slot].OrderSeq:=Buffer.Records[r].SampleSeq;
    Buffer.BatchOwners[Slot].CreatedMs:=Buffer.Records[r].CompletedMonoMs;
    IF NOT windowOpen THEN lastStart:=NowMs; windowOpen:=TRUE; END_IF;
    first:=FALSE; Stage:=10; Busy:=TRUE; ItemPhase:=0;
END_IF;
(* Recheck the same absolute scan deadline before every envelope fragment.
   The dictionary stays pinned by queued records; identity is never read from
   a subsequently changed live configuration. No record is dequeued here. *)
IF Stage=10 THEN
    IF Buffer.WorkDeadlineUs>0 THEN IF GET_MICROSECONDS(TRUE)+ULINT#240>=Buffer.WorkDeadlineUs THEN RETURN; END_IF; END_IF;
    Packets[Slot].Payload:=CONCAT('{"schemaVersion":1,"gatewayId":',NG_Quote(Buffer.Configs[ConfigSlot].GatewayId),',"timestamp":',TO_STRING(HeaderUnixMs,'{0:d}'));
    Stage:=11;
END_IF;
IF Stage=11 THEN
    IF Buffer.WorkDeadlineUs>0 THEN IF GET_MICROSECONDS(TRUE)+ULINT#240>=Buffer.WorkDeadlineUs THEN RETURN; END_IF; END_IF;
    Packets[Slot].Payload:=CONCAT(Packets[Slot].Payload,',"messageId":',NG_Quote(Packets[Slot].MessageId),',"bootId":',NG_Quote(Buffer.Configs[ConfigSlot].CaptureBootId));
    Stage:=12;
END_IF;
IF Stage=12 THEN
    IF Buffer.WorkDeadlineUs>0 THEN IF GET_MICROSECONDS(TRUE)+ULINT#180>=Buffer.WorkDeadlineUs THEN RETURN; END_IF; END_IF;
    Packets[Slot].Payload:=CONCAT(Packets[Slot].Payload,',"sequence":',TO_STRING(HeaderSequence,'{0:d}'),',"configVersion":',TO_STRING(Buffer.Configs[ConfigSlot].Config.Version,'{0:d}'),',"values":[');
    Stage:=1;
END_IF;
IF Stage=1 THEN
    offset:=(Slot-1)*64; finish:=FALSE;
    FOR n:=1 TO 16 DO
        IF Buffer.WorkDeadlineUs=0 THEN IF n>4 THEN EXIT; END_IF;
        ELSIF GET_MICROSECONDS(TRUE)+ULINT#100>=Buffer.WorkDeadlineUs THEN EXIT; END_IF;
        r:=Buffer.QueueHead[Category];
        IF r=0 THEN finish:=TRUE; EXIT; END_IF;
        IF Buffer.Records[r].ConfigSlot<>ConfigSlot THEN finish:=TRUE; EXIT; END_IF;
        pointIndex:=Buffer.Records[r].PointIndex;
        IF (pointIndex<1) OR (pointIndex>320) THEN Buffer.CaptureStopped:=TRUE; RETURN; END_IF;
        (* Epochs replace the growing scan of batch references. This is still
           exact point-index deduplication within one frozen config/batch. *)
        duplicate:=seenPointEpoch[pointIndex]=seenEpoch;
        IF duplicate OR (Buffer.BatchOwners[Slot].Count>=64) OR
           (Buffer.BatchOwners[Slot].Count>=Buffer.Configs[ConfigSlot].Config.maxBatchPoints) THEN finish:=TRUE; EXIT; END_IF;
        (* Until append succeeds the source remains queued. Maintenance may
           expire/reuse its record between slices; never append a stale item. *)
        IF ItemPhase>0 THEN
            IF (ItemRecord<>r) OR (ItemGeneration<>Buffer.RecordGenerations[r]) THEN ItemPhase:=0; END_IF;
        END_IF;
        IF ItemPhase=0 THEN
        IF Buffer.WorkDeadlineUs>0 THEN IF GET_MICROSECONDS(TRUE)+ULINT#180>=Buffer.WorkDeadlineUs THEN EXIT; END_IF; END_IF;
        d:=TO_INT(Buffer.Configs[ConfigSlot].PointDevices[Buffer.Records[r].PointIndex]);
        IF (d>0) AND (d<=Buffer.Configs[ConfigSlot].Config.DeviceCount) THEN
            deviceId:=Buffer.Configs[ConfigSlot].Config.Devices[d].deviceId;
        ELSE
        deviceId:='';
        FOR d:=1 TO Buffer.Configs[ConfigSlot].Config.DeviceCount DO
            IF (Buffer.Records[r].PointIndex>=TO_UINT(Buffer.Configs[ConfigSlot].Config.Devices[d].PointStart)) AND
               (Buffer.Records[r].PointIndex<TO_UINT(Buffer.Configs[ConfigSlot].Config.Devices[d].PointStart+Buffer.Configs[ConfigSlot].Config.Devices[d].PointCount)) THEN
                deviceId:=Buffer.Configs[ConfigSlot].Config.Devices[d].deviceId; EXIT;
            END_IF;
        END_FOR;
            IF deviceId<>'' THEN Buffer.Configs[ConfigSlot].PointDevices[Buffer.Records[r].PointIndex]:=TO_USINT(d); END_IF;
        END_IF;
        valueJson:='null';
        IF Buffer.Records[r].Quality=2 THEN
            IF Buffer.Configs[ConfigSlot].Config.Points[Buffer.Records[r].PointIndex].dataType='bool' THEN
                IF Buffer.Records[r].Value=LREAL#0.0 THEN valueJson:='false'; ELSE valueJson:='true'; END_IF;
            ELSE valueJson:=TO_STRING(Buffer.Records[r].Value,'{0:E16}'); END_IF;
        END_IF;
        IF (d>0) AND (d<=50) THEN
            IF DeviceQuoteSeen[d]<>DeviceQuoteEpoch THEN
                DeviceQuotes[d]:=NG_Quote(deviceId); DeviceQuoteSeen[d]:=DeviceQuoteEpoch;
            END_IF;
            QuotedDevice:=DeviceQuotes[d];
        ELSE QuotedDevice:=NG_Quote(deviceId); END_IF;
        (* Only numeric UTC and quality code determine these text fragments.
           Keys are the original frozen record values, never live time/state. *)
        IF NOT HaveUtc OR (CachedUtc<>Buffer.Records[r].CapturedUtcMs) THEN
            CachedUtc:=Buffer.Records[r].CapturedUtcMs;
            CachedUtcText:=TO_STRING(CachedUtc,'{0:d}'); HaveUtc:=TRUE;
        END_IF;
        IF NOT HaveQuality OR (CachedQuality<>Buffer.Records[r].Quality) THEN
            CachedQuality:=Buffer.Records[r].Quality;
            CachedQualityText:=NG_Quote(NG_QualityName(CachedQuality)); HaveQuality:=TRUE;
        END_IF;
        ItemRecord:=r; ItemGeneration:=Buffer.RecordGenerations[r]; ItemPhase:=1;
        END_IF;
        IF ItemPhase=1 THEN
        IF Buffer.WorkDeadlineUs>0 THEN IF GET_MICROSECONDS(TRUE)+ULINT#180>=Buffer.WorkDeadlineUs THEN EXIT; END_IF; END_IF;
        item:=CONCAT('{"deviceId":',QuotedDevice,',"pointId":',NG_Quote(Buffer.Configs[ConfigSlot].Config.Points[pointIndex].pointId),',"value":',valueJson,',"quality":',CachedQualityText,',"timestamp":',CachedUtcText,'}');
        bytesNeeded:=LEN(Packets[Slot].Payload)+LEN(item)+2;
        IF Buffer.BatchOwners[Slot].Count>0 THEN bytesNeeded:=bytesNeeded+1; END_IF;
        IF bytesNeeded>16380 THEN finish:=TRUE; EXIT; END_IF;
        (* Prefix the small item so the growing full payload is copied once per value. *)
        IF Buffer.BatchOwners[Slot].Count>0 THEN item:=CONCAT(',',item); END_IF;
        ItemPhase:=2;
        END_IF;
        IF Buffer.WorkDeadlineUs>0 THEN IF GET_MICROSECONDS(TRUE)+ULINT#100>=Buffer.WorkDeadlineUs THEN EXIT; END_IF; END_IF;
        Packets[Slot].Payload:=CONCAT(Packets[Slot].Payload,item);
        Buffer.BatchOwners[Slot].Count:=Buffer.BatchOwners[Slot].Count+1; j:=Buffer.BatchOwners[Slot].Count;
        seenPointEpoch[pointIndex]:=seenEpoch;
        Buffer.BatchRefs[offset+j]:=r; Buffer.BatchRefGenerations[offset+j]:=Buffer.RecordGenerations[r];
        Buffer.RecordStates[r]:=2;
        Buffer.QueueHead[Category]:=Buffer.FreeSlots[r]; IF Buffer.QueueHead[Category]=0 THEN Buffer.QueueTail[Category]:=0; END_IF;
        Buffer.FreeSlots[r]:=0;
        ItemPhase:=0;
    END_FOR;
    IF finish THEN
        IF Buffer.BatchOwners[Slot].Count=0 THEN Buffer.CaptureStopped:=TRUE; RETURN; END_IF;
        Packets[Slot].Payload:=CONCAT(Packets[Slot].Payload,']}'); Packets[Slot].Length:=TO_UDINT(LEN(Packets[Slot].Payload)); Stage:=2;
    END_IF;
END_IF;
IF Stage=2 THEN
    Digest(Execute:=TRUE,Length:=Packets[Slot].Length,DeadlineUs:=Buffer.WorkDeadlineUs,Payload:=Packets[Slot].Payload);
    IF Digest.Error THEN Buffer.CaptureStopped:=TRUE; Buffer.AccountingComplete:=FALSE; RETURN; END_IF;
    IF Digest.Done THEN
        IF Buffer.WorkDeadlineUs>0 THEN IF GET_MICROSECONDS(TRUE)+ULINT#100>=Buffer.WorkDeadlineUs THEN RETURN; END_IF; END_IF;
        Buffer.BatchOwners[Slot].Digest:=Digest.Digest; Buffer.BatchOwners[Slot].State:=2;
        Audit(Slot:=Slot,MessageId:=Packets[Slot].MessageId,Buffer:=Buffer);
        Buffer.PreferMaterialize:=TO_USINT(UINT#3-Category); Stage:=0;
    END_IF;
END_IF;
Busy:=Stage<>0;
END_FUNCTION_BLOCK

(* ---- NG_BufferMaintenance.st ---- *)
FUNCTION_BLOCK NG_BufferMaintenance
VAR_INPUT
    GateOpen : BOOL;
    NowMs : ULINT;
END_VAR
VAR_IN_OUT
    Buffer : NG_Buffer;
    Packets : ARRAY[1..16] OF NG_Packet;
END_VAR
VAR
    EndBatch : NG_EndBatch;
    Free : NG_FreeRecord;
    Gap : NG_GapLog;
    Prune : NG_PruneTerminal;
    r : UINT;
    c : UINT;
    q : UINT;
    oldestSlot : UINT;
    oldestSeq : ULINT;
    oldestTerminal : UINT;
    deadSlot : UINT;
    deadCount : UINT;
    deadBytes : UDINT;
    n : INT;
    pressure : BOOL;
    expired : BOOL;
    preparingNew : BOOL;
    stalledNew : BOOL;
    histCount : UINT;
END_VAR
IF Buffer.WorkDeadlineUs>0 THEN IF GET_MICROSECONDS(TRUE)+ULINT#200>=Buffer.WorkDeadlineUs THEN RETURN; END_IF; END_IF;
IF GateOpen AND NOT Buffer.GateWasOpen THEN
    Buffer.Watermark:=Buffer.LastAdmittedSeq;
    IF Buffer.QueueHead[2]<>0 THEN
        IF Buffer.QueueHead[1]=0 THEN Buffer.QueueHead[1]:=Buffer.QueueHead[2];
        ELSE Buffer.FreeSlots[Buffer.QueueTail[1]]:=Buffer.QueueHead[2]; END_IF;
        Buffer.QueueTail[1]:=Buffer.QueueTail[2]; Buffer.QueueHead[2]:=0; Buffer.QueueTail[2]:=0;
    END_IF;
    FOR q:=1 TO 16 DO IF Buffer.BatchOwners[q].State<>0 THEN Buffer.BatchOwners[q].Category:=1; END_IF; END_FOR;
ELSIF GateOpen AND (Buffer.QueueHead[2]<>0) THEN
    (* Hub outage while MQTT stays UP: if live batches stall >=8s without DATA_ACK
       and Queue[2] head ages >=8s, demote aged live records/batches to HISTORY (1)
       so fresh live samples immediately use the reserved Category=2 lane on recovery. *)
    r:=Buffer.QueueHead[2];
    IF (NowMs>Buffer.Records[r].CompletedMonoMs) AND (NowMs>=Buffer.Records[r].CompletedMonoMs+ULINT#8000) THEN
        preparingNew:=FALSE; stalledNew:=FALSE; histCount:=0;
        FOR q:=1 TO 16 DO
            IF Buffer.BatchOwners[q].State<>0 THEN
                IF Buffer.BatchOwners[q].Category=1 THEN histCount:=histCount+1;
                ELSIF Buffer.BatchOwners[q].State=1 THEN preparingNew:=TRUE;
                ELSIF (Buffer.BatchOwners[q].State=2) AND Packets[q].WasSent THEN
                    IF (Packets[q].Attempts>=UDINT#2) OR (NowMs>=Packets[q].RetryAtMs) OR
                       ((NowMs>Packets[q].LastSentMs) AND (NowMs>=Packets[q].LastSentMs+ULINT#8000)) THEN
                        stalledNew:=TRUE;
                    END_IF;
                END_IF;
            END_IF;
        END_FOR;
        IF stalledNew AND NOT preparingNew THEN
            Buffer.Watermark:=Buffer.LastAdmittedSeq;
            IF Buffer.QueueHead[1]=0 THEN Buffer.QueueHead[1]:=Buffer.QueueHead[2];
            ELSE Buffer.FreeSlots[Buffer.QueueTail[1]]:=Buffer.QueueHead[2]; END_IF;
            Buffer.QueueTail[1]:=Buffer.QueueTail[2]; Buffer.QueueHead[2]:=0; Buffer.QueueTail[2]:=0;
            FOR q:=1 TO 16 DO
                IF (histCount<UINT#7) AND (Buffer.BatchOwners[q].State=2) AND (Buffer.BatchOwners[q].Category=2) AND Packets[q].WasSent THEN
                    IF (Packets[q].Attempts>=UDINT#2) OR (NowMs>=Packets[q].RetryAtMs) OR
                       ((NowMs>Packets[q].LastSentMs) AND (NowMs>=Packets[q].LastSentMs+ULINT#8000)) THEN
                        Buffer.BatchOwners[q].Category:=1; histCount:=histCount+1;
                    END_IF;
                END_IF;
            END_FOR;
        END_IF;
    END_IF;
END_IF;
Buffer.GateWasOpen:=GateOpen;
deadCount:=0; deadBytes:=0; deadSlot:=0;
FOR q:=1 TO 16 DO
    IF Buffer.BatchOwners[q].State=3 THEN
        deadCount:=deadCount+1; deadBytes:=deadBytes+Packets[q].Length;
        IF deadSlot=0 THEN deadSlot:=q;
        ELSIF Buffer.BatchOwners[q].OrderSeq<Buffer.BatchOwners[deadSlot].OrderSeq THEN deadSlot:=q; END_IF;
    END_IF;
END_FOR;
IF deadSlot>0 THEN
    IF (deadCount>4) OR (deadBytes>65536) OR (NowMs>=Buffer.BatchOwners[deadSlot].TerminalMs+600000) THEN
        EndBatch(Slot:=deadSlot,Outcome:=USINT#5,Reason:=USINT#0,NowMs:=NowMs,Buffer:=Buffer,Packets:=Packets); RETURN;
    END_IF;
END_IF;
(* At most 64 single-record releases OR one whole batch per scan. Terminal
   evidence shares the same record quota and is reclaimed before live data. *)
FOR n:=1 TO 64 DO
    pressure:=Buffer.OwnedCount+TO_UDINT(MIN(Buffer.IngressCount,UINT#64))>UDINT#28800;
    IF pressure THEN
        oldestTerminal:=0;
        FOR q:=1 TO 64 DO
            IF Buffer.TerminalOwners[q].Count>0 THEN
                IF oldestTerminal=0 THEN oldestTerminal:=q;
                ELSIF Buffer.TerminalOwners[q].FirstSeq<Buffer.TerminalOwners[oldestTerminal].FirstSeq THEN oldestTerminal:=q; END_IF;
            END_IF;
        END_FOR;
        IF oldestTerminal>0 THEN Prune(Index:=oldestTerminal,Buffer:=Buffer); RETURN; END_IF;
    END_IF;
    c:=0; r:=0; oldestSlot:=0; oldestSeq:=ULINT#9007199254740991;
    FOR q:=1 TO 2 DO
        IF Buffer.QueueHead[q]>0 THEN
            IF Buffer.Records[Buffer.QueueHead[q]].SampleSeq<oldestSeq THEN
                c:=q; r:=Buffer.QueueHead[q]; oldestSeq:=Buffer.Records[r].SampleSeq;
            END_IF;
        END_IF;
    END_FOR;
    FOR q:=1 TO 16 DO
        IF Buffer.BatchOwners[q].State>=2 THEN
            IF Buffer.BatchOwners[q].OrderSeq<oldestSeq THEN oldestSlot:=q; oldestSeq:=Buffer.BatchOwners[q].OrderSeq; r:=0; END_IF;
        END_IF;
    END_FOR;
    expired:=FALSE;
    IF r>0 THEN expired:=NowMs>=Buffer.Records[r].CompletedMonoMs+900000;
    ELSIF oldestSlot>0 THEN expired:=NowMs>=Buffer.BatchOwners[oldestSlot].CreatedMs+900000; END_IF;
    IF NOT pressure AND NOT expired THEN EXIT; END_IF;
    IF r>0 THEN
        Buffer.QueueHead[c]:=Buffer.FreeSlots[r]; IF Buffer.QueueHead[c]=0 THEN Buffer.QueueTail[c]:=0; END_IF;
        Buffer.KnownUnsentEventsTotal:=NG_SafeAdd(Buffer.KnownUnsentEventsTotal,ULINT#1);
        IF expired THEN Gap(Reason:=USINT#6,Event:=Buffer.Records[r],Buffer:=Buffer); ELSE Gap(Reason:=USINT#5,Event:=Buffer.Records[r],Buffer:=Buffer); END_IF;
        Free(Index:=r,Buffer:=Buffer);
    ELSIF oldestSlot>0 THEN
        q:=2; IF Packets[oldestSlot].WasSent THEN q:=4; END_IF;
        IF Buffer.BatchOwners[oldestSlot].State=3 THEN q:=5; END_IF;
        c:=5; IF expired THEN c:=6; END_IF;
        EndBatch(Slot:=oldestSlot,Outcome:=TO_USINT(q),Reason:=TO_USINT(c),NowMs:=NowMs,Buffer:=Buffer,Packets:=Packets);
        (* Under a hard full-pool fence even terminal evidence must yield to
           new capture. Preserve the cumulative U/I fact and gap, explicitly
           mark evidence pruning rather than reject a fresh cohort silently. *)
        IF pressure AND (q>=4) THEN Prune(Index:=Buffer.TerminalIndex,Buffer:=Buffer); END_IF;
        RETURN;
    ELSE EXIT; END_IF;
END_FOR;
END_FUNCTION_BLOCK

(* ---- NG_Capture.st ---- *)
FUNCTION_BLOCK NG_Capture
VAR_INPUT
    PointIndex : UINT;
    Kind : USINT;
    Quality : USINT;
    Value : LREAL;
    NowMs : ULINT;
    NominalDueMs : ULINT;
    SystemUtcMs : ULINT;
END_VAR
VAR_OUTPUT
    Accepted : BOOL;
END_VAR
VAR_IN_OUT
    Buffer : NG_Buffer;
END_VAR
VAR
    Core : NG_CaptureCore;
END_VAR
(* Validate the index before binding the cursor reference. *)
Accepted:=FALSE;
IF Buffer.CaptureStopped OR NOT Buffer.LayoutValid OR (Buffer.ActiveSlot=0) OR (Buffer.ActiveSlot>4) THEN RETURN; END_IF;
IF (PointIndex<1) OR (PointIndex>320) THEN Buffer.CaptureStopped:=TRUE; RETURN; END_IF;
Core(PointIndex:=PointIndex,Kind:=Kind,Quality:=Quality,Value:=Value,NowMs:=NowMs,NominalDueMs:=NominalDueMs,SystemUtcMs:=SystemUtcMs,Cursor:=Buffer.Cursors[PointIndex],Buffer:=Buffer);
Accepted:=Core.Accepted;
END_FUNCTION_BLOCK

(* ---- NG_CaptureCore.st ---- *)
FUNCTION_BLOCK NG_CaptureCore
VAR_INPUT
    PointIndex : UINT;
    Kind : USINT;
    Quality : USINT;
    Value : LREAL;
    NowMs : ULINT;
    NominalDueMs : ULINT;
    SystemUtcMs : ULINT;
END_VAR
VAR_OUTPUT
    Accepted : BOOL;
END_VAR
VAR_IN_OUT
    Cursor : NG_SourceCursor;
    Buffer : NG_Buffer;
END_VAR
VAR
    s : UINT;
    d : INT;
    Gap : NG_GapLog;
    Audit : NG_AuditCapture;
    AuditDecision : NG_AuditDecision;
END_VAR

Accepted:=FALSE; s:=Buffer.ActiveSlot;
IF Buffer.CaptureStopped OR NOT Buffer.LayoutValid OR (s=0) OR (s>4) THEN RETURN; END_IF;
IF (PointIndex<1) OR (PointIndex>320) THEN Buffer.CaptureStopped:=TRUE; RETURN; END_IF;
IF (Buffer.NextSampleSeq>=ULINT#9007199254740991) OR (NowMs>ULINT#9007199254740991) THEN
    Buffer.CaptureStopped:=TRUE; RETURN;
END_IF;
Buffer.NextSampleSeq:=Buffer.NextSampleSeq+1;
Buffer.CapturedEventsTotal:=NG_SafeAdd(Buffer.CapturedEventsTotal,ULINT#1);
Buffer.Scratch.SampleSeq:=Buffer.NextSampleSeq; Buffer.Scratch.Value:=0;
IF Quality=2 THEN Buffer.Scratch.Value:=Value; END_IF;
Buffer.Scratch.Kind:=Kind; Buffer.Scratch.Quality:=Quality;
Buffer.Scratch.CompletedMonoMs:=NowMs; Buffer.Scratch.NominalDueMonoMs:=0;
Buffer.Scratch.ConfigSlot:=s; Buffer.Scratch.ConfigGeneration:=Buffer.Configs[s].Generation;
Buffer.Scratch.PointIndex:=PointIndex; Buffer.Scratch.SamplingGeneration:=Buffer.SamplingGeneration;
Buffer.Scratch.ClockRevision:=0; Buffer.Scratch.CapturedUtcMs:=0; Buffer.Scratch.Flags:=WORD#8;
(* Explicit SYSTEM_RTC_COMPAT_UNVERIFIED: trusted UTC/timeValid remain absent. *)
IF (SystemUtcMs>0) AND (SystemUtcMs<=ULINT#9007199254740991) THEN Buffer.Scratch.CapturedUtcMs:=SystemUtcMs; Buffer.Scratch.Flags:=WORD#9; END_IF;
IF Buffer.PlatformTime THEN
    Buffer.Scratch.ClockRevision:=Buffer.ClockRevision; Buffer.Scratch.CapturedUtcMs:=0; Buffer.Scratch.Flags:=WORD#0;
    IF Buffer.TimeValid AND (SystemUtcMs>0) AND (SystemUtcMs<=ULINT#9007199254740991) THEN
        Buffer.Scratch.CapturedUtcMs:=SystemUtcMs; Buffer.Scratch.Flags:=WORD#3;
    END_IF;
END_IF;
IF Kind=1 THEN
    Buffer.Scratch.NominalDueMonoMs:=NominalDueMs; Buffer.Scratch.Flags:=Buffer.Scratch.Flags OR WORD#4;
    IF Cursor.HasPhysicalUtc AND ((Buffer.Scratch.Flags AND WORD#1)<>WORD#0) AND
       (Cursor.LastPhysicalUtcMs=SystemUtcMs) THEN
        Buffer.SourceTimestampRepeatTotal:=NG_SafeAdd(Buffer.SourceTimestampRepeatTotal,ULINT#1);
    END_IF;
    Cursor.HasPhysicalUtc:=(Buffer.Scratch.Flags AND WORD#1)<>WORD#0;
    Cursor.LastPhysicalUtcMs:=SystemUtcMs;
END_IF;
Audit(Buffer:=Buffer,Event:=Buffer.Scratch);
IF Buffer.IngressCount>=512 THEN
    Buffer.CaptureOverflowEventsTotal:=NG_SafeAdd(Buffer.CaptureOverflowEventsTotal,ULINT#1);
    Buffer.AccountingComplete:=FALSE;
    Buffer.UndecidedLostEventsTotal:=NG_SafeAdd(Buffer.UndecidedLostEventsTotal,ULINT#1);
    Gap(Reason:=USINT#1,Outcome:=USINT#5,Event:=Buffer.Scratch,Buffer:=Buffer);
    AuditDecision(SampleSeq:=Buffer.Scratch.SampleSeq,Decision:=USINT#4,Reason:=USINT#1,Buffer:=Buffer);
    RETURN;
END_IF;
Buffer.Ingress[Buffer.Tail]:=Buffer.Scratch; Buffer.Tail:=Buffer.Tail MOD 512+1;
Buffer.IngressCount:=Buffer.IngressCount+1; Buffer.Configs[s].References:=Buffer.Configs[s].References+1;
Accepted:=TRUE;
END_FUNCTION_BLOCK

(* ---- NG_Char.st ---- *)
FUNCTION_BLOCK NG_Char
VAR_INPUT
    Code : UDINT;
    Utf8 : BOOL;
END_VAR
VAR_OUTPUT
    Value : STRING[4];
END_VAR
VAR
    Bytes : ARRAY[0..4] OF BYTE;
    Convert : BUF_TO_STRING;
    Count : INT;
END_VAR
Count := 1;
Bytes[0] := TO_BYTE(Code);
IF Utf8 THEN
    IF Code < 128 THEN Bytes[0] := TO_BYTE(Code);
    ELSIF Code < 2048 THEN Count := 2; Bytes[0] := TO_BYTE(192 + Code / 64); Bytes[1] := TO_BYTE(128 + Code MOD 64);
    ELSIF Code < 65536 THEN Count := 3; Bytes[0] := TO_BYTE(224 + Code / 4096); Bytes[1] := TO_BYTE(128 + (Code / 64) MOD 64); Bytes[2] := TO_BYTE(128 + Code MOD 64);
    ELSE Count := 4; Bytes[0] := TO_BYTE(240 + Code / 262144); Bytes[1] := TO_BYTE(128 + (Code / 4096) MOD 64); Bytes[2] := TO_BYTE(128 + (Code / 64) MOD 64); Bytes[3] := TO_BYTE(128 + Code MOD 64);
    END_IF;
END_IF;
Bytes[Count] := BYTE#0;
Convert(REQ := FALSE, BUF_FORMAT := FALSE, BUF_OFFS := 0, BUF_CNT := Count, BUFFER := Bytes, DST := Value);
Convert(REQ := TRUE, BUF_FORMAT := FALSE, BUF_OFFS := 0, BUF_CNT := Count, BUFFER := Bytes, DST := Value);
END_FUNCTION_BLOCK

(* ---- NG_CheckCounters.st ---- *)
FUNCTION_BLOCK NG_CheckCounters
VAR_IN_OUT
    Buffer : NG_Buffer;
END_VAR
VAR
    maximum : ULINT := ULINT#9007199254740991;
END_VAR
IF (Buffer.CapturedEventsTotal>=maximum) OR (Buffer.EligibleEventsTotal>=maximum) OR
   (Buffer.PolicyFilteredEventsTotal>=maximum) OR (Buffer.TimeInvalidEventsTotal>=maximum) OR
   (Buffer.CaptureOverflowEventsTotal>=maximum) OR (Buffer.UndecidedLostEventsTotal>=maximum) OR
   (Buffer.KnownUnsentEventsTotal>=maximum) OR (Buffer.IsolatedEventsTotal>=maximum) OR
   (Buffer.UncertainDeliveryEventsTotal>=maximum) OR (Buffer.StoredConfirmedEventsTotal>=maximum) OR
   (Buffer.LateStoredEventsTotal>=maximum) OR (Buffer.EnqueueRejectedAttemptsTotal>=maximum) OR
   (Buffer.MissedPollCyclesTotal>=maximum) OR (Buffer.MissedReportSlotsTotal>=maximum) OR
   (Buffer.SourceTimestampRepeatTotal>=maximum) OR (Buffer.GapRecordsTotal>=maximum) THEN
    Buffer.CounterOverflow:=TRUE;
END_IF;
IF Buffer.CounterOverflow OR Buffer.CaptureStopped OR (Buffer.UndecidedLostEventsTotal>0) THEN Buffer.AccountingComplete:=FALSE; END_IF;
END_FUNCTION_BLOCK

(* ---- NG_Command.st ---- *)
FUNCTION_BLOCK NG_Command
VAR_INPUT
    Execute : BOOL;
    IsPatch : BOOL;
    Retained : BOOL;
    GatewayId : NG_Id;
END_VAR
VAR_IN_OUT
    Doc : NG_Document;
    Active : NG_Config;
END_VAR
VAR_OUTPUT
    Done : BOOL;
    Candidate : NG_Config;
    ErrorCode : NG_Text;
    RequestId : NG_Id;
    RequestVersion : ULINT;
END_VAR
VAR
    ReadConfig : NG_ReadConfig;
    ReadDevice : NG_ReadDevice;
    Change : NG_EditDevice;
    NewDevice : NG_Device;
    NewPoints : ARRAY[1..32] OF NG_Point;
    Prev : BOOL;
    n : INT;
    t : INT;
    a : INT;
    g : INT;
    r : INT;
    op : INT;
    dev : INT;
    d : INT;
    i : INT;
    count : INT;
    id : NG_Id;
    mode : STRING[16];
    seen : ARRAY[1..50] OF NG_Id;
END_VAR
IF NOT Execute THEN Done := FALSE; Prev := FALSE; RETURN; END_IF;
IF Prev THEN RETURN; END_IF;
Prev := TRUE; Done := TRUE; ErrorCode := 'SCHEMA_INVALID'; RequestId := ''; RequestVersion := 0;
IF IsPatch THEN
    IF NOT NG_Allowed(1,'|schemaVersion|gatewayId|timestamp|messageId|configVersion|baseConfigVersion|baseMessageId|operations|gateway|',Doc) THEN RETURN; END_IF;
ELSE
    IF NOT NG_Allowed(1,'|schemaVersion|gatewayId|timestamp|messageId|configVersion|config|',Doc) THEN RETURN; END_IF;
END_IF;
t := NG_Member(1,'messageId',Doc);
IF (Doc.Tokens[t].Kind <> 3) OR (LEN(Doc.Tokens[t].Text)>64) THEN RETURN; END_IF;
RequestId := Doc.Tokens[t].Text;
IF NOT NG_ValidId(RequestId) THEN RequestId := ''; RETURN; END_IF;
t := NG_Member(1,'configVersion',Doc);
IF (Doc.Tokens[t].Kind <> 4) OR (Doc.Tokens[t].Number < 1) OR (Doc.Tokens[t].Number > LREAL#9007199254740991.0) OR (Doc.Tokens[t].Number <> TO_LREAL(TO_LINT(Doc.Tokens[t].Number))) THEN RETURN; END_IF;
RequestVersion := TO_ULINT(Doc.Tokens[t].Number);
t := NG_Member(1,'schemaVersion',Doc);
IF (Doc.Tokens[t].Kind <> 4) OR (Doc.Tokens[t].Number <> 1) THEN RETURN; END_IF;
t := NG_Member(1,'gatewayId',Doc);
IF (Doc.Tokens[t].Kind <> 3) OR (Doc.Tokens[t].Text <> GatewayId) THEN ErrorCode := 'GATEWAY_MISMATCH'; RETURN; END_IF;
t := NG_Member(1,'timestamp',Doc);
IF (Doc.Tokens[t].Kind <> 4) OR (Doc.Tokens[t].Number < 0) OR (Doc.Tokens[t].Number > LREAL#9007199254740991.0) OR (Doc.Tokens[t].Number <> TO_LREAL(TO_LINT(Doc.Tokens[t].Number))) THEN RETURN; END_IF;
(* Version/replay checks run before this FB in the coordinator. *)
IF NOT IsPatch THEN
    n := NG_Member(1,'config',Doc);
    ReadConfig(Node := n, Doc := Doc, Config := Candidate);
    ErrorCode := ReadConfig.ErrorText;
ELSE
    IF Retained THEN ErrorCode := 'RETAINED_PATCH'; RETURN; END_IF;
    t := NG_Member(1,'baseConfigVersion',Doc);
    IF (Doc.Tokens[t].Kind <> 4) OR (Doc.Tokens[t].Number <> TO_LREAL(Active.Version)) THEN ErrorCode := 'BASE_CONFIG_MISMATCH'; RETURN; END_IF;
    t := NG_Member(1,'baseMessageId',Doc);
    IF Active.Version = 0 THEN
        IF Doc.Tokens[t].Kind <> 6 THEN ErrorCode := 'BASE_CONFIG_MISMATCH'; RETURN; END_IF;
    ELSIF (Doc.Tokens[t].Kind <> 3) OR (Doc.Tokens[t].Text <> Active.MessageId) THEN ErrorCode := 'BASE_CONFIG_MISMATCH'; RETURN;
    END_IF;
    IF RequestVersion <= Active.Version THEN ErrorCode := 'STALE_VERSION'; RETURN; END_IF;
    Candidate := Active;
    g := NG_Member(1,'gateway',Doc);
    IF g > 0 THEN
        IF NOT NG_Allowed(g,'|enabled|report|',Doc) THEN RETURN; END_IF;
        t := NG_Member(g,'enabled',Doc);
        IF t > 0 THEN
            IF Doc.Tokens[t].Kind <> 5 THEN RETURN; END_IF;
            Candidate.enabled := Doc.Tokens[t].Text = 'true';
        ELSIF Active.Version = 0 THEN RETURN; END_IF;
        r := NG_Member(g,'report',Doc);
        IF r > 0 THEN
            IF NOT NG_Allowed(r,'|batchIntervalMs|maxBatchPoints|',Doc) THEN RETURN; END_IF;
            t := NG_Member(r,'batchIntervalMs',Doc);
            IF (Doc.Tokens[t].Kind <> 4) OR (Doc.Tokens[t].Number < 1) OR (Doc.Tokens[t].Number > 86400000) OR (Doc.Tokens[t].Number <> TO_LREAL(TO_LINT(Doc.Tokens[t].Number))) THEN RETURN; END_IF;
            Candidate.batchIntervalMs := TO_UDINT(Doc.Tokens[t].Number);
            t := NG_Member(r,'maxBatchPoints',Doc);
            IF (Doc.Tokens[t].Kind <> 4) OR (Doc.Tokens[t].Number < 1) OR (Doc.Tokens[t].Number > 500) OR (Doc.Tokens[t].Number <> TO_LREAL(TO_LINT(Doc.Tokens[t].Number))) THEN RETURN; END_IF;
            Candidate.maxBatchPoints := TO_UINT(Doc.Tokens[t].Number);
        ELSIF Active.Version = 0 THEN RETURN; END_IF;
    ELSIF Active.Version = 0 THEN RETURN;
    END_IF;
    a := NG_Member(1,'operations',Doc);
    IF Doc.Tokens[a].Kind <> 2 THEN RETURN; END_IF;
    IF (Doc.Tokens[a].NextToken = a+1) AND ((g = 0) OR (Doc.Tokens[g].NextToken = g+1)) THEN RETURN; END_IF;
    op := a+1; count := 0;
    WHILE op < Doc.Tokens[a].NextToken DO
        IF count >= 50 THEN ErrorCode := 'POINT_LIMIT_EXCEEDED'; RETURN; END_IF;
        IF NOT NG_Allowed(op,'|op|deviceId|device|',Doc) THEN RETURN; END_IF;
        t := NG_Member(op,'deviceId',Doc);
        IF (Doc.Tokens[t].Kind <> 3) OR (LEN(Doc.Tokens[t].Text)>64) THEN RETURN; END_IF;
        id := Doc.Tokens[t].Text;
        IF NOT NG_ValidId(id) THEN RETURN; END_IF;
        FOR i := 1 TO count DO IF seen[i] = id THEN ErrorCode := 'OPERATION_CONFLICT'; RETURN; END_IF; END_FOR;
        count := count+1; seen[count] := id;
        t := NG_Member(op,'op',Doc);
        IF Doc.Tokens[t].Kind <> 3 THEN RETURN; END_IF;
        mode := Doc.Tokens[t].Text; d := 0;
        FOR i := 1 TO Candidate.DeviceCount DO IF Candidate.Devices[i].deviceId = id THEN d := i; EXIT; END_IF; END_FOR;
        IF mode = 'add' THEN
            IF d > 0 THEN ErrorCode := 'DEVICE_EXISTS'; RETURN; END_IF;
            IF Candidate.DeviceCount >= 50 THEN ErrorCode := 'POINT_LIMIT_EXCEEDED'; RETURN; END_IF;
            d := Candidate.DeviceCount+1;
        ELSIF (mode = 'replace') OR (mode = 'remove') THEN
            IF d = 0 THEN ErrorCode := 'DEVICE_NOT_FOUND'; RETURN; END_IF;
        ELSE RETURN; END_IF;
        dev := NG_Member(op,'device',Doc);
        IF mode = 'remove' THEN
            IF dev <> 0 THEN RETURN; END_IF;
            Change(DeviceIndex := d, Remove := TRUE, Replacement := NewDevice, Config := Candidate, Points := NewPoints);
            IF Change.ErrorText <> '' THEN ErrorCode := Change.ErrorText; RETURN; END_IF;
        ELSE
            ReadDevice(Node := dev, Doc := Doc, Device := NewDevice, Points := NewPoints);
            ErrorCode := ReadDevice.ErrorText;
            IF ErrorCode <> '' THEN RETURN; END_IF;
            ErrorCode := 'SCHEMA_INVALID';
            IF NewDevice.deviceId <> id THEN ErrorCode := 'OPERATION_CONFLICT'; RETURN; END_IF;
        END_IF;
        IF mode <> 'remove' THEN
            Change(DeviceIndex := d, Remove := FALSE, Replacement := NewDevice, Config := Candidate, Points := NewPoints);
            IF Change.ErrorText <> '' THEN ErrorCode := Change.ErrorText; RETURN; END_IF;
        END_IF;
        op := Doc.Tokens[op].NextToken;
    END_WHILE;
    ErrorCode := NG_CheckConfig(Candidate);
END_IF;
Candidate.Version := RequestVersion; Candidate.MessageId := RequestId;
END_FUNCTION_BLOCK

(* ---- NG_ConfigSlot.st ---- *)
FUNCTION_BLOCK NG_ConfigSlot
VAR_INPUT
    GatewayId : NG_Id;
    CaptureBootId : NG_Id;
END_VAR
VAR_OUTPUT
    Slot : UINT;
END_VAR
VAR_IN_OUT
    Config : NG_Config;
    Buffer : NG_Buffer;
END_VAR
VAR
    Compare : NG_SameConfig;
    Prune : NG_PruneTerminal;
    i : INT;
    j : INT;
    oldIndex : UINT;
    configSlot : UINT;
    recIndex : UINT;
    hasFree : BOOL;
END_VAR
Slot := 0;
IF Buffer.ActiveSlot>0 THEN
    Compare(A:=Buffer.Configs[Buffer.ActiveSlot].Config,B:=Config);
    IF (Buffer.Configs[Buffer.ActiveSlot].GatewayId=GatewayId) AND
       (Buffer.Configs[Buffer.ActiveSlot].CaptureBootId=CaptureBootId) AND
       Compare.Equal THEN
        Slot:=Buffer.ActiveSlot; RETURN;
    END_IF;
END_IF;
IF Buffer.NextConfigGeneration=UDINT#4294967295 THEN Buffer.CaptureStopped:=TRUE; RETURN; END_IF;
FOR i:=1 TO 4 DO
    IF (i<>TO_INT(Buffer.ActiveSlot)) AND (Buffer.Configs[i].References=0) AND NOT Buffer.Configs[i].Reserved THEN
        Buffer.NextConfigGeneration:=Buffer.NextConfigGeneration+1;
        Buffer.Configs[i].Config:=Config; Buffer.Configs[i].GatewayId:=GatewayId;
        Buffer.Configs[i].CaptureBootId:=CaptureBootId;
        Buffer.Configs[i].Generation:=Buffer.NextConfigGeneration;
        FOR j:=1 TO 320 DO Buffer.Configs[i].PointDevices[j]:=0; END_FOR;
        Buffer.Configs[i].Reserved:=TRUE; Slot:=TO_UINT(i); RETURN;
    END_IF;
END_FOR;
(* When no external audit collector is attached, evict oldest audit/association
   ring entries on dictionary exhaustion so inactive config slots can be freed
   without dropping live Ingress/Records/Outbox telemetry. *)
IF (Buffer.AuditAckBootId<>CaptureBootId) AND (Buffer.AssociationAckBootId<>CaptureBootId) THEN
    hasFree:=FALSE;
    WHILE (NOT hasFree) AND (Buffer.AuditReadSeq<Buffer.AuditWriteSeq) DO
        oldIndex:=TO_UINT(Buffer.AuditReadSeq MOD 512)+1;
        configSlot:=Buffer.AuditEvents[oldIndex].Event.ConfigSlot;
        IF (configSlot<1) OR (configSlot>4) THEN Buffer.CaptureStopped:=TRUE; Buffer.EvidenceComplete:=FALSE; RETURN; END_IF;
        IF Buffer.Configs[configSlot].References=0 THEN Buffer.CaptureStopped:=TRUE; Buffer.EvidenceComplete:=FALSE; RETURN; END_IF;
        Buffer.Configs[configSlot].References:=Buffer.Configs[configSlot].References-1;
        Buffer.AuditReadSeq:=Buffer.AuditReadSeq+1;
        Buffer.AuditDropped:=NG_SafeAdd(Buffer.AuditDropped,ULINT#1);
        Buffer.EvidenceComplete:=FALSE;
        IF (configSlot<>Buffer.ActiveSlot) AND (Buffer.Configs[configSlot].References=0) AND NOT Buffer.Configs[configSlot].Reserved THEN
            hasFree:=TRUE;
        END_IF;
    END_WHILE;
    WHILE (NOT hasFree) AND (Buffer.AssociationReadSeq<Buffer.AssociationWriteSeq) DO
        oldIndex:=TO_UINT(Buffer.AssociationReadSeq MOD 32)+1;
        configSlot:=Buffer.Associations[oldIndex].ConfigSlot;
        IF (configSlot<1) OR (configSlot>4) THEN Buffer.CaptureStopped:=TRUE; Buffer.EvidenceComplete:=FALSE; RETURN; END_IF;
        IF Buffer.Configs[configSlot].References=0 THEN Buffer.CaptureStopped:=TRUE; Buffer.EvidenceComplete:=FALSE; RETURN; END_IF;
        Buffer.Configs[configSlot].References:=Buffer.Configs[configSlot].References-1;
        Buffer.AssociationReadSeq:=Buffer.AssociationReadSeq+1;
        Buffer.AssociationDropped:=NG_SafeAdd(Buffer.AssociationDropped,ULINT#1);
        Buffer.EvidenceComplete:=FALSE;
        IF (configSlot<>Buffer.ActiveSlot) AND (Buffer.Configs[configSlot].References=0) AND NOT Buffer.Configs[configSlot].Reserved THEN
            hasFree:=TRUE;
        END_IF;
    END_WHILE;
    IF NOT hasFree THEN
        FOR i:=1 TO 64 DO
            IF Buffer.TerminalOwners[i].Count>0 THEN
                recIndex:=Buffer.TerminalRefs[(i-1)*64+1];
                IF (recIndex>0) AND (recIndex<=Buffer.HighSlot) THEN
                    configSlot:=Buffer.Records[recIndex].ConfigSlot;
                    IF (configSlot>=1) AND (configSlot<=4) AND (configSlot<>Buffer.ActiveSlot) THEN
                        Prune(Index:=TO_UINT(i),Buffer:=Buffer);
                        IF (Buffer.Configs[configSlot].References=0) AND NOT Buffer.Configs[configSlot].Reserved THEN
                            hasFree:=TRUE; EXIT;
                        END_IF;
                    END_IF;
                END_IF;
            END_IF;
        END_FOR;
    END_IF;
    FOR i:=1 TO 4 DO
        IF (i<>TO_INT(Buffer.ActiveSlot)) AND (Buffer.Configs[i].References=0) AND NOT Buffer.Configs[i].Reserved THEN
            Buffer.NextConfigGeneration:=Buffer.NextConfigGeneration+1;
            Buffer.Configs[i].Config:=Config; Buffer.Configs[i].GatewayId:=GatewayId;
            Buffer.Configs[i].CaptureBootId:=CaptureBootId;
            Buffer.Configs[i].Generation:=Buffer.NextConfigGeneration;
            FOR j:=1 TO 320 DO Buffer.Configs[i].PointDevices[j]:=0; END_FOR;
            Buffer.Configs[i].Reserved:=TRUE; Slot:=TO_UINT(i); RETURN;
        END_IF;
    END_FOR;
END_IF;
END_FUNCTION_BLOCK

(* ---- NG_Delivery.st ---- *)
FUNCTION_BLOCK NG_Delivery
VAR_INPUT
    GateOpen : BOOL;
    NowMs : ULINT;
    GatewayId : NG_Id;
    BootId : NG_Id;
    SubmitAck : BOOL;
    AckMessageId : NG_Id;
    AckStored : BOOL;
    AckRetryable : BOOL;
    AckCodes : NG_Text;
END_VAR
VAR_IN_OUT
    Buffer : NG_Buffer;
    Packets : ARRAY[1..16] OF NG_Packet;
END_VAR
VAR_OUTPUT
    AckBusy : BOOL;
    SendSlot : UINT;
    SendGeneration : UDINT;
    SendMessageId : NG_Id;
END_VAR
VAR
    Digest : NG_StringSHA256;
    EndBatch : NG_EndBatch;
    Free : NG_FreeRecord;
    pendingAck : BOOL;
    ackId : NG_Id;
    stored : BOOL;
    retryable : BOOL;
    codes : NG_Text;
    op : UINT; (* 1 verify send,2 verify ACK *)
    slot : UINT;
    generation : UDINT;
    id : NG_Id;
    q : UINT;
    j : UINT;
    r : UINT;
    c : UINT;
    terminal : UINT;
    inFlight : UINT;
    inHistory : UINT;
    inNew : UINT;
    candidates : ARRAY[1..2] OF UINT;
    offset : UINT;
    valid : BOOL;
    eligible : BOOL;
END_VAR
IF SubmitAck AND NOT pendingAck THEN
    pendingAck:=TRUE; ackId:=AckMessageId; stored:=AckStored; retryable:=AckRetryable; codes:=AckCodes;
    IF op=1 THEN op:=0; SendSlot:=0; END_IF;
END_IF;
AckBusy:=pendingAck OR (op=2);
IF SendSlot>0 THEN
    IF NOT GateOpen OR (Buffer.BatchGenerations[SendSlot]<>SendGeneration) OR
       (Buffer.BatchOwners[SendSlot].State<>2) OR (Packets[SendSlot].MessageId<>SendMessageId) OR
       (NowMs<Packets[SendSlot].RetryAtMs) THEN SendSlot:=0; END_IF;
END_IF;
IF op<>0 THEN
    IF (Buffer.BatchGenerations[slot]<>generation) OR (Packets[slot].MessageId<>id) OR (Buffer.BatchOwners[slot].State<2) THEN
        IF op=2 THEN pendingAck:=FALSE; END_IF;
        op:=0;
    END_IF;
END_IF;
IF op=0 THEN
    IF Buffer.WorkDeadlineUs>0 THEN IF GET_MICROSECONDS(TRUE)+ULINT#180>=Buffer.WorkDeadlineUs THEN RETURN; END_IF; END_IF;
    Digest(Execute:=FALSE,Length:=UDINT#0,Payload:=Packets[1].Payload);
    IF pendingAck THEN
        SendSlot:=0; slot:=0;
        FOR q:=1 TO 16 DO
            IF (Packets[q].MessageId=ackId) AND (Buffer.BatchOwners[q].State>=2) AND Packets[q].WasSent THEN slot:=q; EXIT; END_IF;
        END_FOR;
        IF slot>0 THEN
            generation:=Buffer.BatchGenerations[slot]; id:=ackId; op:=2;
        ELSE
            terminal:=0;
            FOR q:=1 TO 64 DO
                IF (Buffer.TerminalOwners[q].Count>0) AND (Buffer.TerminalOwners[q].MessageId=ackId) THEN terminal:=q; EXIT; END_IF;
            END_FOR;
            IF terminal=0 THEN Buffer.UnknownAcksTotal:=NG_SafeAdd(Buffer.UnknownAcksTotal,ULINT#1);
            ELSIF stored THEN
                IF Buffer.TerminalOwners[terminal].Outcome=2 THEN Buffer.ConflictingAcksTotal:=NG_SafeAdd(Buffer.ConflictingAcksTotal,ULINT#1);
                ELSE
                    offset:=(terminal-1)*64; valid:=Buffer.TerminalOwners[terminal].Digest<>'';
                    FOR j:=1 TO Buffer.TerminalOwners[terminal].Count DO
                        r:=Buffer.TerminalRefs[offset+j];
                        IF r=0 THEN valid:=FALSE;
                        ELSIF (Buffer.RecordGenerations[r]<>Buffer.TerminalRefGenerations[offset+j]) OR (Buffer.RecordStates[r]<>3) THEN valid:=FALSE;
                        ELSIF (Buffer.Configs[Buffer.Records[r].ConfigSlot].GatewayId<>GatewayId) OR
                              (Buffer.Configs[Buffer.Records[r].ConfigSlot].CaptureBootId<>BootId) THEN valid:=FALSE; END_IF;
                    END_FOR;
                    IF valid THEN
                        FOR j:=1 TO Buffer.TerminalOwners[terminal].Count DO
                            r:=Buffer.TerminalRefs[offset+j]; Free(Index:=r,Buffer:=Buffer);
                            Buffer.StoredConfirmedEventsTotal:=NG_SafeAdd(Buffer.StoredConfirmedEventsTotal,ULINT#1);
                            Buffer.LateStoredEventsTotal:=NG_SafeAdd(Buffer.LateStoredEventsTotal,ULINT#1);
                            Buffer.TerminalRefs[offset+j]:=0;
                        END_FOR;
                        Buffer.TerminalOwners[terminal].Count:=0; Buffer.TerminalOwners[terminal].Outcome:=3;
                    ELSE Buffer.CaptureStopped:=TRUE; END_IF;
                END_IF;
            END_IF;
            pendingAck:=FALSE;
        END_IF;
    (* Verify during the pacing wait; actual submission still gates NextSendAt. *)
    ELSIF GateOpen AND (SendSlot=0) THEN
        inFlight:=0; inHistory:=0; inNew:=0; candidates[1]:=0; candidates[2]:=0;
        FOR q:=1 TO 16 DO
            IF (Buffer.BatchOwners[q].State=2) AND Packets[q].WasSent THEN
                inFlight:=inFlight+1;
                IF Buffer.BatchOwners[q].Category=1 THEN inHistory:=inHistory+1; ELSE inNew:=inNew+1; END_IF;
            END_IF;
        END_FOR;
        FOR q:=1 TO 16 DO
            IF Buffer.BatchOwners[q].State=2 THEN
                c:=TO_UINT(Buffer.BatchOwners[q].Category);
                IF (c<1) OR (c>2) THEN Buffer.CaptureStopped:=TRUE; Buffer.AccountingComplete:=FALSE; RETURN; END_IF;
                eligible:=Packets[q].WasSent OR ((inFlight<8) AND (((c=1) AND (inHistory<7)) OR ((c=2) AND (inNew<7))));
                eligible:=eligible AND (NowMs>=Packets[q].RetryAtMs);
                IF eligible THEN
                    IF candidates[c]=0 THEN candidates[c]:=q;
                    ELSIF Buffer.BatchOwners[q].OrderSeq<Buffer.BatchOwners[candidates[c]].OrderSeq THEN candidates[c]:=q; END_IF;
                END_IF;
            END_IF;
        END_FOR;
        c:=TO_UINT(Buffer.PreferSend); IF candidates[c]=0 THEN c:=UINT#3-c; END_IF;
        slot:=candidates[c];
        IF slot>0 THEN generation:=Buffer.BatchGenerations[slot]; id:=Packets[slot].MessageId; op:=1; END_IF;
    END_IF;
END_IF;
IF op<>0 THEN
    Digest(Execute:=TRUE,Length:=Packets[slot].Length,DeadlineUs:=Buffer.WorkDeadlineUs,Payload:=Packets[slot].Payload);
    IF Digest.Error THEN Buffer.CaptureStopped:=TRUE; Buffer.AccountingComplete:=FALSE; RETURN; END_IF;
    IF Digest.Done THEN
        IF Buffer.WorkDeadlineUs>0 THEN IF GET_MICROSECONDS(TRUE)+ULINT#350>=Buffer.WorkDeadlineUs THEN RETURN; END_IF; END_IF;
        valid:=(Digest.Digest=Buffer.BatchOwners[slot].Digest) AND (Packets[slot].Length=TO_UDINT(LEN(Packets[slot].Payload)));
        c:=Buffer.BatchOwners[slot].ConfigSlot;
        IF (c<1) OR (c>4) THEN Buffer.CaptureStopped:=TRUE; Buffer.AccountingComplete:=FALSE; op:=0; pendingAck:=FALSE; RETURN; END_IF;
        valid:=valid AND (Buffer.Configs[c].GatewayId=GatewayId) AND (Buffer.Configs[c].CaptureBootId=BootId);
        offset:=(slot-1)*64;
        FOR j:=1 TO Buffer.BatchOwners[slot].Count DO
            r:=Buffer.BatchRefs[offset+j];
            IF r=0 THEN valid:=FALSE;
            ELSIF Buffer.RecordGenerations[r]<>Buffer.BatchRefGenerations[offset+j] THEN valid:=FALSE; END_IF;
        END_FOR;
        IF NOT valid THEN
            Buffer.CorruptBatchesTotal:=NG_SafeAdd(Buffer.CorruptBatchesTotal,ULINT#1); Buffer.CaptureStopped:=TRUE;
            Buffer.AccountingComplete:=FALSE;
            IF Buffer.BatchOwners[slot].State=2 THEN
                c:=2; IF Packets[slot].WasSent THEN c:=4; END_IF;
                EndBatch(Slot:=slot,Outcome:=TO_USINT(c),Reason:=USINT#7,NowMs:=NowMs,Buffer:=Buffer,Packets:=Packets);
            END_IF;
        ELSIF op=2 THEN
            IF stored THEN
                IF Buffer.BatchOwners[slot].State=3 THEN Buffer.ConflictingAcksTotal:=NG_SafeAdd(Buffer.ConflictingAcksTotal,ULINT#1);
                ELSE EndBatch(Slot:=slot,Outcome:=USINT#1,Reason:=USINT#0,NowMs:=NowMs,Buffer:=Buffer,Packets:=Packets); END_IF;
            ELSIF Buffer.BatchOwners[slot].State=2 THEN
                IF retryable THEN Packets[slot].RetryAtMs:=MAX(Packets[slot].RetryAtMs,NowMs+60000+TO_ULINT(slot)*17); Packets[slot].LastError:=codes;
                ELSE Packets[slot].LastError:=codes; EndBatch(Slot:=slot,Outcome:=USINT#3,Reason:=USINT#8,NowMs:=NowMs,Buffer:=Buffer,Packets:=Packets); END_IF;
            END_IF;
        ELSIF GateOpen AND (NowMs>=Packets[slot].RetryAtMs) THEN
            SendSlot:=slot; SendGeneration:=generation; SendMessageId:=id;
        END_IF;
        IF op=2 THEN pendingAck:=FALSE; END_IF;
        op:=0;
    END_IF;
END_IF;
AckBusy:=pendingAck OR (op=2);
END_FUNCTION_BLOCK

(* ---- NG_DeliveryParallel.st ---- *)
FUNCTION_BLOCK NG_DeliveryParallel
VAR_INPUT
    GateOpen : BOOL;
    NowMs : ULINT;
    GatewayId : NG_Id;
    BootId : NG_Id;
    SubmitAck : BOOL;
    AckMessageId : NG_Id;
    AckStored : BOOL;
    AckRetryable : BOOL;
    AckCodes : NG_Text;
END_VAR
VAR_IN_OUT
    Buffer : NG_Buffer;
    Packets : ARRAY[1..16] OF NG_Packet;
END_VAR
VAR_OUTPUT
    AckBusy : BOOL;
    SendSlot : UINT;
    SendGeneration : UDINT;
    SendMessageId : NG_Id;
END_VAR
VAR
    AckPath : NG_Delivery;
    SendPath : NG_Delivery;
    preferAck : BOOL;
    priorityHold : BOOL;
END_VAR
(* Independent bounded hash state prevents an incoming ACK from repeatedly
   cancelling an unfinished send verification. Both paths keep the original
   immutable SHA-256 and generation checks; ACK is serialised first. *)
(* Main rotates builder/delivery every scan. Flipping this priority every scan
   locks both clocks together: send always wins the delivery-first scans.
   Hold each inner priority for two calls, giving ACK and send one full-budget
   delivery-first turn each in every four scans. Neither digest is restarted. *)
priorityHold:=NOT priorityHold;
IF priorityHold THEN preferAck:=NOT preferAck; END_IF;
IF preferAck THEN
AckPath(GateOpen:=FALSE,NowMs:=NowMs,GatewayId:=GatewayId,BootId:=BootId,SubmitAck:=SubmitAck,
    AckMessageId:=AckMessageId,AckStored:=AckStored,AckRetryable:=AckRetryable,AckCodes:=AckCodes,Buffer:=Buffer,Packets:=Packets);
SendPath(GateOpen:=GateOpen,NowMs:=NowMs,GatewayId:=GatewayId,BootId:=BootId,SubmitAck:=FALSE,
    AckMessageId:='',AckStored:=FALSE,AckRetryable:=FALSE,AckCodes:='',Buffer:=Buffer,Packets:=Packets);
ELSE
SendPath(GateOpen:=GateOpen,NowMs:=NowMs,GatewayId:=GatewayId,BootId:=BootId,SubmitAck:=FALSE,
    AckMessageId:='',AckStored:=FALSE,AckRetryable:=FALSE,AckCodes:='',Buffer:=Buffer,Packets:=Packets);
AckPath(GateOpen:=FALSE,NowMs:=NowMs,GatewayId:=GatewayId,BootId:=BootId,SubmitAck:=SubmitAck,
    AckMessageId:=AckMessageId,AckStored:=AckStored,AckRetryable:=AckRetryable,AckCodes:=AckCodes,Buffer:=Buffer,Packets:=Packets);
END_IF;
AckBusy:=AckPath.AckBusy; SendSlot:=SendPath.SendSlot; SendGeneration:=SendPath.SendGeneration; SendMessageId:=SendPath.SendMessageId;
END_FUNCTION_BLOCK

(* ---- NG_Diagnostics.st ---- *)
FUNCTION_BLOCK NG_Diagnostics
VAR_INPUT
    BootId : NG_Id;
    GatewayId : NG_Id;
    NowMs : ULINT;
    Force : BOOL;
END_VAR
VAR_IN_OUT
    Buffer : NG_Buffer;
END_VAR
VAR
    lastUpdate : ULINT;
    oldest : ULINT;
    hasOldest : BOOL;
    q : UINT;
    r : UINT;
    pendingBatches : UINT;
    deadBatches : UINT;
END_VAR
IF NOT Buffer.DiagnosticInitialized THEN
    Buffer.DiagnosticInitialized:=TRUE;
    Buffer.RestartLossUnknown:=TRUE; Buffer.AccountingComplete:=FALSE;
    Buffer.GapRecordsTotal:=NG_SafeAdd(Buffer.GapRecordsTotal,ULINT#1);
    Buffer.Diagnostics.LastGap.Reason:=9; Buffer.Diagnostics.LastGap.Outcome:=4;
    Buffer.Diagnostics.LastGapCountKnown:=FALSE;
END_IF;
IF NOT Force AND (NowMs<lastUpdate+1000) AND (Buffer.Diagnostics.Revision<>0) THEN RETURN; END_IF;
IF NOT Force AND (Buffer.WorkDeadlineUs>0) THEN IF GET_MICROSECONDS(TRUE)+ULINT#350>=Buffer.WorkDeadlineUs THEN RETURN; END_IF; END_IF;
IF Buffer.Diagnostics.Revision>=ULINT#9007199254740988 THEN Buffer.CounterOverflow:=TRUE; RETURN; END_IF;
Buffer.Diagnostics.Revision:=Buffer.Diagnostics.Revision+1;
Buffer.Diagnostics.BootId:=BootId; Buffer.Diagnostics.GatewayId:=GatewayId;
Buffer.Diagnostics.CapturedMonoMs:=NowMs;
IF Buffer.ActiveSlot>0 THEN Buffer.Diagnostics.ConfigVersion:=Buffer.Configs[Buffer.ActiveSlot].Config.Version; END_IF;
Buffer.Diagnostics.Totals[1]:=Buffer.CapturedEventsTotal;
Buffer.Diagnostics.Totals[2]:=Buffer.EligibleEventsTotal;
Buffer.Diagnostics.Totals[3]:=Buffer.PolicyFilteredEventsTotal;
Buffer.Diagnostics.Totals[4]:=Buffer.TimeInvalidEventsTotal;
Buffer.Diagnostics.Totals[5]:=Buffer.CaptureOverflowEventsTotal;
Buffer.Diagnostics.Totals[6]:=Buffer.UndecidedLostEventsTotal;
Buffer.Diagnostics.Totals[7]:=Buffer.KnownUnsentEventsTotal;
Buffer.Diagnostics.Totals[8]:=Buffer.IsolatedEventsTotal;
Buffer.Diagnostics.Totals[9]:=Buffer.UncertainDeliveryEventsTotal;
Buffer.Diagnostics.Totals[10]:=Buffer.StoredConfirmedEventsTotal;
Buffer.Diagnostics.Totals[11]:=Buffer.LateStoredEventsTotal;
Buffer.Diagnostics.Totals[12]:=Buffer.EnqueueRejectedAttemptsTotal;
Buffer.Diagnostics.Totals[13]:=Buffer.MissedPollCyclesTotal;
Buffer.Diagnostics.Totals[14]:=Buffer.MissedReportSlotsTotal;
Buffer.Diagnostics.Totals[15]:=Buffer.SourceTimestampRepeatTotal;
Buffer.Diagnostics.Totals[16]:=Buffer.GapRecordsTotal;
Buffer.Diagnostics.DecisionPending:=TO_ULINT(Buffer.IngressCount);
Buffer.Diagnostics.PendingEvents:=TO_ULINT(Buffer.OwnedCount)-Buffer.DeadRetainedEvents-Buffer.UncertainRetainedEvents+TO_ULINT(Buffer.IngressCount);
Buffer.Diagnostics.DeadEvents:=Buffer.DeadRetainedEvents;
Buffer.Diagnostics.UncertainRetainedEvents:=Buffer.UncertainRetainedEvents;
oldest:=ULINT#9007199254740991; hasOldest:=FALSE; pendingBatches:=0; deadBatches:=0;
IF Buffer.IngressCount>0 THEN oldest:=Buffer.Ingress[Buffer.Head].CompletedMonoMs; hasOldest:=TRUE; END_IF;
FOR q:=1 TO 2 DO
    r:=Buffer.QueueHead[q];
    IF r>0 THEN oldest:=MIN(oldest,Buffer.Records[r].CompletedMonoMs); hasOldest:=TRUE; END_IF;
END_FOR;
FOR q:=1 TO 16 DO
    IF Buffer.BatchOwners[q].State=2 THEN pendingBatches:=pendingBatches+1; END_IF;
    IF Buffer.BatchOwners[q].State=3 THEN deadBatches:=deadBatches+1; END_IF;
    IF (Buffer.BatchOwners[q].State=1) OR (Buffer.BatchOwners[q].State=2) THEN oldest:=MIN(oldest,Buffer.BatchOwners[q].CreatedMs); hasOldest:=TRUE; END_IF;
END_FOR;
Buffer.Diagnostics.PendingBatches:=pendingBatches; Buffer.Diagnostics.DeadBatches:=deadBatches;
Buffer.Diagnostics.OldestPendingAgeMs:=0; Buffer.Diagnostics.HasPendingAge:=FALSE;
IF hasOldest AND (NowMs>=oldest) THEN Buffer.Diagnostics.OldestPendingAgeMs:=NowMs-oldest; Buffer.Diagnostics.HasPendingAge:=TRUE; END_IF;
Buffer.Diagnostics.AllocatedBytes:=Buffer.LayoutBytes;
Buffer.Diagnostics.UsedBytes:=Buffer.LayoutBytes-(UDINT#28800-Buffer.OwnedCount)*Buffer.RecordBytes;
Buffer.Diagnostics.MaxBytes:=4194304;
Buffer.Diagnostics.AccountingComplete:=Buffer.AccountingComplete;
Buffer.Diagnostics.CounterOverflow:=Buffer.CounterOverflow; Buffer.Diagnostics.DetailTruncated:=Buffer.DetailTruncated;
Buffer.Diagnostics.RestartLossUnknown:=Buffer.RestartLossUnknown;
Buffer.Diagnostics.AuditDropped:=Buffer.AuditDropped; Buffer.Diagnostics.AssociationDropped:=Buffer.AssociationDropped;
Buffer.Diagnostics.EvidenceComplete:=Buffer.EvidenceComplete;
IF Buffer.GapIndex>0 THEN Buffer.Diagnostics.LastGap:=Buffer.Gaps[Buffer.GapIndex]; Buffer.Diagnostics.LastGapCountKnown:=TRUE; END_IF;
Buffer.Diagnostics.HmiSummary:=CONCAT('RAM P=',TO_STRING(Buffer.Diagnostics.PendingEvents,'{0:d}'),' I=',TO_STRING(Buffer.Diagnostics.DeadEvents,'{0:d}'),' U-retained=',TO_STRING(Buffer.Diagnostics.UncertainRetainedEvents,'{0:d}'),' bytes=',TO_STRING(Buffer.Diagnostics.UsedBytes,'{0:d}'),'/',TO_STRING(Buffer.Diagnostics.MaxBytes,'{0:d}'),' restart-loss=UNKNOWN auditDrops=',TO_STRING(Buffer.AuditDropped+Buffer.AssociationDropped,'{0:d}'));
Buffer.Diagnostics.Revision:=Buffer.Diagnostics.Revision+1; lastUpdate:=NowMs;
END_FUNCTION_BLOCK

(* ---- NG_EditDevice.st ---- *)
FUNCTION_BLOCK NG_EditDevice
VAR_INPUT
    DeviceIndex : INT;
    Remove : BOOL;
    Replacement : NG_Device;
END_VAR
VAR_IN_OUT
    Config : NG_Config;
    Points : ARRAY[1..32] OF NG_Point;
END_VAR
VAR_OUTPUT
    ErrorText : NG_Text;
END_VAR
VAR
    oldCount : INT;
    newCount : INT;
    start : INT;
    delta : INT;
    i : INT;
    n : INT;
END_VAR
ErrorText := 'SCHEMA_INVALID';
IF (DeviceIndex < 1) OR (DeviceIndex > Config.DeviceCount+1) OR (DeviceIndex > 50) THEN RETURN; END_IF;
oldCount := 0; start := Config.PointCount+1;
IF DeviceIndex <= Config.DeviceCount THEN oldCount := Config.Devices[DeviceIndex].PointCount; start := Config.Devices[DeviceIndex].PointStart; END_IF;
newCount := Replacement.PointCount; IF Remove THEN newCount := 0; END_IF;
delta := newCount-oldCount;
IF (newCount < 0) OR (newCount > 32) OR (Config.PointCount+delta > 320) THEN ErrorText := 'POINT_LIMIT_EXCEEDED'; RETURN; END_IF;
IF delta > 0 THEN
    FOR i := Config.PointCount TO start+oldCount BY -1 DO Config.Points[i+delta] := Config.Points[i]; END_FOR;
ELSIF delta < 0 THEN
    FOR i := start+oldCount TO Config.PointCount DO Config.Points[i+delta] := Config.Points[i]; END_FOR;
END_IF;
Config.PointCount := Config.PointCount+delta;
IF Remove THEN
    IF DeviceIndex > Config.DeviceCount THEN RETURN; END_IF;
    FOR i := DeviceIndex TO Config.DeviceCount-1 DO Config.Devices[i] := Config.Devices[i+1]; END_FOR;
    Config.DeviceCount := Config.DeviceCount-1;
ELSE
    Config.Devices[DeviceIndex] := Replacement;
    IF DeviceIndex > Config.DeviceCount THEN Config.DeviceCount := DeviceIndex; END_IF;
    FOR i := 1 TO newCount DO Config.Points[start+i-1] := Points[i]; END_FOR;
END_IF;
n := 1;
FOR i := 1 TO Config.DeviceCount DO Config.Devices[i].PointStart := n; n := n+Config.Devices[i].PointCount; END_FOR;
ErrorText := '';
END_FUNCTION_BLOCK

(* ---- NG_EndBatch.st ---- *)
FUNCTION_BLOCK NG_EndBatch
VAR_INPUT
    Slot : UINT;
    Outcome : USINT; (* 1 STORED,2 known unsent,3 permanent isolated,4 uncertain,5 prune isolated *)
    Reason : USINT;
    NowMs : ULINT;
END_VAR
VAR_IN_OUT
    Buffer : NG_Buffer;
    Packets : ARRAY[1..16] OF NG_Packet;
END_VAR
VAR
    Free : NG_FreeRecord;
    Gap : NG_GapLog;
    Prune : NG_PruneTerminal;
    j : UINT;
    r : UINT;
    offset : UINT;
    terminalOffset : UINT;
    terminal : UINT;
END_VAR
IF (Slot=0) OR (Slot>16) THEN RETURN; END_IF;
IF Buffer.BatchOwners[Slot].State<2 THEN RETURN; END_IF;
IF (Outcome=3) AND (Buffer.BatchOwners[Slot].State=3) THEN RETURN; END_IF;
offset:=(Slot-1)*64; terminal:=0;
(* Validate the whole ownership set before any irreversible counter/release. *)
FOR j:=1 TO Buffer.BatchOwners[Slot].Count DO
    r:=Buffer.BatchRefs[offset+j];
    IF r=0 THEN Buffer.CaptureStopped:=TRUE; Buffer.AccountingComplete:=FALSE; RETURN; END_IF;
    IF (Buffer.RecordGenerations[r]<>Buffer.BatchRefGenerations[offset+j]) OR (Buffer.RecordStates[r]=0) THEN
        Buffer.CaptureStopped:=TRUE; Buffer.AccountingComplete:=FALSE; RETURN;
    END_IF;
END_FOR;
IF Outcome=1 THEN Buffer.StoredBatchesTotal:=NG_SafeAdd(Buffer.StoredBatchesTotal,ULINT#1); END_IF;
IF (Outcome=4) OR (Outcome=5) THEN
    Buffer.TerminalIndex:=Buffer.TerminalIndex MOD 64+1; terminal:=Buffer.TerminalIndex;
    Prune(Index:=terminal,Buffer:=Buffer); terminalOffset:=(terminal-1)*64;
    Buffer.TerminalOwners[terminal].MessageId:=Packets[Slot].MessageId;
    Buffer.TerminalOwners[terminal].Digest:=Buffer.BatchOwners[Slot].Digest;
    Buffer.TerminalOwners[terminal].BatchGeneration:=Buffer.BatchGenerations[Slot];
    Buffer.TerminalOwners[terminal].Count:=Buffer.BatchOwners[Slot].Count;
    Buffer.TerminalOwners[terminal].FirstSeq:=Buffer.BatchOwners[Slot].OrderSeq;
    Buffer.TerminalOwners[terminal].CreatedMs:=NowMs;
    Buffer.TerminalOwners[terminal].Outcome:=1;
    IF Outcome=5 THEN Buffer.TerminalOwners[terminal].Outcome:=2;
        Buffer.DeadPrunedBatchesTotal:=NG_SafeAdd(Buffer.DeadPrunedBatchesTotal,ULINT#1); END_IF;
END_IF;
FOR j:=1 TO Buffer.BatchOwners[Slot].Count DO
    r:=Buffer.BatchRefs[offset+j];
    IF (r=0) OR (Buffer.RecordGenerations[r]<>Buffer.BatchRefGenerations[offset+j]) THEN Buffer.CaptureStopped:=TRUE; RETURN; END_IF;
    CASE Outcome OF
    1: Buffer.StoredConfirmedEventsTotal:=NG_SafeAdd(Buffer.StoredConfirmedEventsTotal,ULINT#1); Free(Index:=r,Buffer:=Buffer);
    2: Buffer.KnownUnsentEventsTotal:=NG_SafeAdd(Buffer.KnownUnsentEventsTotal,ULINT#1); Gap(Reason:=Reason,Outcome:=USINT#2,Event:=Buffer.Records[r],Buffer:=Buffer); Free(Index:=r,Buffer:=Buffer);
    3: Buffer.IsolatedEventsTotal:=NG_SafeAdd(Buffer.IsolatedEventsTotal,ULINT#1); Gap(Reason:=Reason,Outcome:=USINT#3,Event:=Buffer.Records[r],Buffer:=Buffer); Buffer.RecordStates[r]:=4; Buffer.DeadRetainedEvents:=Buffer.DeadRetainedEvents+1;
    4: Buffer.UncertainDeliveryEventsTotal:=NG_SafeAdd(Buffer.UncertainDeliveryEventsTotal,ULINT#1); Gap(Reason:=Reason,Outcome:=USINT#4,Event:=Buffer.Records[r],Buffer:=Buffer); Buffer.RecordStates[r]:=3; Buffer.UncertainRetainedEvents:=Buffer.UncertainRetainedEvents+1;
    END_CASE;
    IF terminal>0 THEN
        Buffer.TerminalRefs[terminalOffset+j]:=r;
        Buffer.TerminalRefGenerations[terminalOffset+j]:=Buffer.RecordGenerations[r];
    END_IF;
    IF Outcome<>3 THEN Buffer.BatchRefs[offset+j]:=0; END_IF;
END_FOR;
IF Outcome=3 THEN
    Buffer.BatchOwners[Slot].State:=3; Buffer.BatchOwners[Slot].TerminalMs:=NowMs; Packets[Slot].Dead:=TRUE;
ELSE
    Buffer.BatchOwners[Slot].State:=0; Buffer.BatchOwners[Slot].Count:=0;
    Packets[Slot].MessageId:=''; Packets[Slot].Payload:=''; Packets[Slot].Length:=0;
    Packets[Slot].WasSent:=FALSE; Packets[Slot].Dead:=FALSE; Packets[Slot].Attempts:=0;
    Packets[Slot].LastSentMs:=0; Packets[Slot].RetryAtMs:=0; Packets[Slot].LastError:='';
END_IF;
END_FUNCTION_BLOCK

(* ---- NG_FreeRecord.st ---- *)
FUNCTION_BLOCK NG_FreeRecord
VAR_INPUT
    Index : UINT;
END_VAR
VAR_IN_OUT
    Buffer : NG_Buffer;
END_VAR
VAR
    s : UINT;
END_VAR
IF (Index=0) OR (Index>Buffer.HighSlot) THEN RETURN; END_IF;
IF Buffer.RecordStates[Index]=0 THEN Buffer.CaptureStopped:=TRUE; RETURN; END_IF;
s:=Buffer.Records[Index].ConfigSlot;
IF Buffer.Configs[s].References=0 THEN Buffer.CaptureStopped:=TRUE; RETURN; END_IF;
Buffer.Configs[s].References:=Buffer.Configs[s].References-1;
IF Buffer.RecordStates[Index]=4 THEN Buffer.DeadRetainedEvents:=Buffer.DeadRetainedEvents-1; END_IF;
IF Buffer.RecordStates[Index]=3 THEN Buffer.UncertainRetainedEvents:=Buffer.UncertainRetainedEvents-1; END_IF;
Buffer.RecordStates[Index]:=0; Buffer.FreeSlots[Index]:=Buffer.FreeHead;
Buffer.FreeHead:=Index; Buffer.OwnedCount:=Buffer.OwnedCount-1;
END_FUNCTION_BLOCK

(* ---- NG_GapLog.st ---- *)
FUNCTION_BLOCK NG_GapLog
VAR_INPUT
    Reason : USINT; (* 1 overflow,2 version,4 time,5 capacity,6 age,7 corrupt *)
    Outcome : USINT;
END_VAR
VAR_IN_OUT
    Event : NG_CaptureEvent;
    Buffer : NG_Buffer;
END_VAR
VAR
    s : UINT;
    p : UINT;
    d : INT;
END_VAR
s:=Event.ConfigSlot; p:=Event.PointIndex;
Buffer.GapRecordsTotal:=NG_SafeAdd(Buffer.GapRecordsTotal,ULINT#1);
Buffer.GapIndex:=Buffer.GapIndex MOD 64+1;
IF Buffer.GapRecordsTotal>64 THEN Buffer.DetailTruncated:=TRUE; END_IF;
Buffer.Gaps[Buffer.GapIndex].SampleSeq:=Event.SampleSeq;
Buffer.Gaps[Buffer.GapIndex].CompletedMonoMs:=Event.CompletedMonoMs;
Buffer.Gaps[Buffer.GapIndex].Reason:=Reason;
Buffer.Gaps[Buffer.GapIndex].Outcome:=Outcome;
IF Outcome=0 THEN
    Buffer.Gaps[Buffer.GapIndex].Outcome:=2;
    IF (Reason=1) OR (Reason=2) THEN Buffer.Gaps[Buffer.GapIndex].Outcome:=5; END_IF;
END_IF;
Buffer.Gaps[Buffer.GapIndex].CapturedUtcMs:=Event.CapturedUtcMs;
Buffer.Gaps[Buffer.GapIndex].Flags:=Event.Flags;
Buffer.Gaps[Buffer.GapIndex].ConfigVersion:=Buffer.Configs[s].Config.Version;
Buffer.Gaps[Buffer.GapIndex].GatewayId:=Buffer.Configs[s].GatewayId;
Buffer.Gaps[Buffer.GapIndex].CaptureBootId:=Buffer.Configs[s].CaptureBootId;
Buffer.Gaps[Buffer.GapIndex].PointId:=Buffer.Configs[s].Config.Points[p].pointId;
Buffer.Gaps[Buffer.GapIndex].DeviceId:='';
FOR d:=1 TO Buffer.Configs[s].Config.DeviceCount DO
    IF (p>=TO_UINT(Buffer.Configs[s].Config.Devices[d].PointStart)) AND
       (p<TO_UINT(Buffer.Configs[s].Config.Devices[d].PointStart+Buffer.Configs[s].Config.Devices[d].PointCount)) THEN
        Buffer.Gaps[Buffer.GapIndex].DeviceId:=Buffer.Configs[s].Config.Devices[d].deviceId; EXIT;
    END_IF;
END_FOR;
END_FUNCTION_BLOCK
